(* IEC 61131-3 sources: PortalRobot/Portal_robot/Device/application, 34 files *)

(* ---- Persistent_Value.gvl.st ---- *)
{attribute 'qualified_only'}
VAR_GLOBAL PERSISTENT RETAIN
	// Постоянное хранилище базовых точек в энергонезависимой памяти контроллера.
	// Размер 15 сохранён ради совместимости со старой раскладкой: позиции 2, 6 и 10
	// (legacy MACHINE_x_INSIDE) больше не публикуются и не участвуют в готовности.
	astRetainPoints : ARRAY [1..GVL_POINT.iPersistentPointCapacity] OF ST_POINT;
	udiPointStorageVersion : UDINT;

	// Геометрический контроль: настройки, память станций и вызовы.
	astConfig : ARRAY [1..2] OF ST_GEOMETRY_CONFIG;
	astMemory : ARRAY [1..2] OF ST_GEOMETRY_MEMORY;
	astRetainCalls : ARRAY [1..3] OF ST_GEOMETRY_CALL;
	udiNextCallId : UDINT;
	udiEventSequence : UDINT;
	xAutoEnabled : BOOL := FALSE;
	auiPeriod : ARRAY [1..3] OF UINT := [20, 20, 20];
	auiCount : ARRAY [1..3] OF UINT;
	xWaitWhenOccupied : BOOL := TRUE;
	tTransportTimeout : TIME := T#10S;
	tDriveFeedbackTimeout : TIME := T#3S;
	tResetPulse : TIME := T#1S;
	tWaitWarningTimeout : TIME := T#180S; // Ожидание готовой вызванной детали в станке до WARNING

	// Постоянный шаг сетки для расчёта координат робота, отдельно по типам магазинов.
	lrStaticPitchX : LREAL := 60.0;
	lrStaticPitchY : LREAL := 60.0;
	lrTwinPitchX : LREAL := 70.0;
	lrTwinPitchY : LREAL := 70.0;

	// Базы ГК для SIMULATION сохраняются отдельно от реальных координат.
	astSimulationConfig : ARRAY [1..2] OF ST_GEOMETRY_CONFIG;

	// Добавлено в конце списка: прежние 15 баз и их версия сохраняют раскладку.
	astMagazineCalibration : ARRAY [1..2] OF ST_MAGAZINE_CALIBRATION;
END_VAR

(* ---- PLC_PRG.AppendIoEvent.st ---- *)
METHOD PRIVATE AppendIoEvent
VAR_INPUT
    usiDirection : USINT;
    uiIndex : UINT;
    usiKind : USINT;
    xOld : BOOL;
    xNew : BOOL;
END_VAR
VAR
    uiSlot : UINT;
    sEvent : STRING(96);
END_VAR

// --- BEGIN IMPLEMENTATION ---

IF NOT xIoSnapshotPublishing THEN
    GVL_HMI.udiIoJournalRevision := GVL_HMI.udiIoJournalRevision + UDINT#1;
END_IF;
// Переполнение Seq открывает новый FIFO; идентификаторы не повторяются внутри эпохи.
IF GVL_HMI.udiIoJournalSequence = UDINT#4294967295 THEN
    GVL_HMI.udiIoBootCounter := GVL_HMI.udiIoBootCounter + UDINT#1;
    IF GVL_HMI.udiIoBootCounter = UDINT#0 THEN GVL_HMI.udiIoBootCounter := UDINT#1; END_IF;
    GVL_HMI.udiIoJournalSequence := UDINT#0;
    GVL_HMI.uiIoJournalHead := UINT#0;
    GVL_HMI.uiIoJournalCount := UINT#0;
END_IF;
uiSlot := (GVL_HMI.uiIoJournalHead MOD UINT#100) + UINT#1;
GVL_HMI.udiIoJournalSequence := GVL_HMI.udiIoJournalSequence + UDINT#1;
astIoEvent[uiSlot].udiSequence := GVL_HMI.udiIoJournalSequence;
astIoEvent[uiSlot].uliTimeMs := uliIoClockMs;
astIoEvent[uiSlot].usiDirection := usiDirection;
astIoEvent[uiSlot].uiIndex := uiIndex;
astIoEvent[uiSlot].usiKind := usiKind;
astIoEvent[uiSlot].xOld := xOld;
astIoEvent[uiSlot].xNew := xNew;
// Строка кодируется только для изменившегося слота, не для всего FIFO на каждом скане.
sEvent := CONCAT(UDINT_TO_STRING(GVL_HMI.udiIoJournalSequence), ';');
sEvent := CONCAT(sEvent, ULINT_TO_STRING(uliIoClockMs));
sEvent := CONCAT(sEvent, ';'); sEvent := CONCAT(sEvent, USINT_TO_STRING(usiDirection));
sEvent := CONCAT(sEvent, ';'); sEvent := CONCAT(sEvent, UINT_TO_STRING(uiIndex));
sEvent := CONCAT(sEvent, ';'); sEvent := CONCAT(sEvent, USINT_TO_STRING(usiKind));
sEvent := CONCAT(sEvent, ';'); sEvent := CONCAT(sEvent, USINT_TO_STRING(BOOL_TO_USINT(xOld)));
sEvent := CONCAT(sEvent, ';'); sEvent := CONCAT(sEvent, USINT_TO_STRING(BOOL_TO_USINT(xNew)));
GVL_HMI.asIoJournal[uiSlot] := sEvent;
GVL_HMI.uiIoJournalHead := uiSlot;
GVL_HMI.uiIoJournalCount := MIN(UINT#100, GVL_HMI.uiIoJournalCount + UINT#1);
IF NOT xIoSnapshotPublishing THEN
    GVL_HMI.udiIoJournalRevision := GVL_HMI.udiIoJournalRevision + UDINT#1;
END_IF;

(* ---- PLC_PRG.ApplyIoOutputOverrides.st ---- *)
METHOD PRIVATE ApplyIoOutputOverrides

// --- BEGIN IMPLEMENTATION ---

// Прямой ручной режим владеет всеми DO. Штатные уровни остаются отдельно для возврата программе.
axIoAutoDo[1] := GVL_PHYSICAL_IO.xDoMachine1HatchClosed;
axIoAutoDo[2] := GVL_PHYSICAL_IO.xDoMachine1HatchUnLock;
axIoAutoDo[3] := GVL_PHYSICAL_IO.xDoMachine1ClampChuck;
axIoAutoDo[4] := GVL_PHYSICAL_IO.xDoMachine1UnclampChuck;
axIoAutoDo[5] := GVL_PHYSICAL_IO.xDoMachine1StartCycle;
axIoAutoDo[6] := GVL_PHYSICAL_IO.xDoMachine2HatchClosed;
axIoAutoDo[7] := GVL_PHYSICAL_IO.xDoMachine2HatchUnLock;
axIoAutoDo[8] := GVL_PHYSICAL_IO.xDoMachine2ClampChuck;
axIoAutoDo[9] := GVL_PHYSICAL_IO.xDoMachine2UnclampChuck;
axIoAutoDo[10] := GVL_PHYSICAL_IO.xDoMachine2StartCycle;
axIoAutoDo[11] := GVL_PHYSICAL_IO.xDoMachine3HatchClosed;
axIoAutoDo[12] := GVL_PHYSICAL_IO.xDoMachine3HatchUnLock;
axIoAutoDo[13] := GVL_PHYSICAL_IO.xDoMachine3ClampChuck;
axIoAutoDo[14] := GVL_PHYSICAL_IO.xDoMachine3UnclampChuck;
axIoAutoDo[15] := GVL_PHYSICAL_IO.xDoMachine3StartCycle;
axIoAutoDo[16] := GVL_PHYSICAL_IO.xDoGripper1Open;
axIoAutoDo[17] := GVL_PHYSICAL_IO.xDoGripper2Open;
axIoAutoDo[18] := GVL_PHYSICAL_IO.xDoRotateToDetail;
axIoAutoDo[19] := GVL_PHYSICAL_IO.xDoDoor1Unlock;
axIoAutoDo[20] := GVL_PHYSICAL_IO.xDoDoor2Unlock;
axIoAutoDo[21] := GVL_PHYSICAL_IO.xDoDoor3Unlock;
axIoAutoDo[22] := GVL_PHYSICAL_IO.xDoDoor4Unlock;
axIoAutoDo[23] := GVL_PHYSICAL_IO.xDoSafetyRelayReset;
axIoAutoDo[24] := GVL_PHYSICAL_IO.xDoSignalTowerGreenOutput;
axIoAutoDo[25] := GVL_PHYSICAL_IO.xDoSignalTowerAmberOutput;
axIoAutoDo[26] := GVL_PHYSICAL_IO.xDoSignalTowerRedOutput;
axIoAutoDo[27] := GVL_PHYSICAL_IO.xDoDoor1ButtonLamp;
axIoAutoDo[28] := GVL_PHYSICAL_IO.xDoDoor2ButtonLamp;
axIoAutoDo[29] := GVL_PHYSICAL_IO.xDoDoor3ButtonLamp;
axIoAutoDo[30] := GVL_PHYSICAL_IO.xDoDoor4ButtonLamp;
axIoAutoDo[31] := GVL_PHYSICAL_IO.xDoMagazine1LockIn;
axIoAutoDo[32] := GVL_PHYSICAL_IO.xDoMagazine1LockOut;
axIoAutoDo[33] := GVL_PHYSICAL_IO.xDoMagazine1StopIn;
axIoAutoDo[34] := GVL_PHYSICAL_IO.xDoMagazine1StopOut;
axIoAutoDo[35] := GVL_PHYSICAL_IO.xDoMagazine1LiftUp;
axIoAutoDo[36] := GVL_PHYSICAL_IO.xDoMagazine1LiftDown;
axIoAutoDo[37] := FALSE; // Удалённый сигнал; индекс журнала не переиспользовать.
axIoAutoDo[38] := FALSE; // Удалённый сигнал; индекс журнала не переиспользовать.
axIoAutoDo[39] := FALSE; // Удалённый сигнал; индекс журнала не переиспользовать.
axIoAutoDo[40] := GVL_PHYSICAL_IO.xDoCellAlarmHorn;
axIoAutoDo[41] := GVL_PHYSICAL_IO.xDoGk1DriveRun;
axIoAutoDo[42] := GVL_PHYSICAL_IO.xDoGk1DriveReset;
axIoAutoDo[43] := GVL_PHYSICAL_IO.xDoMagazine2LockIn;
axIoAutoDo[44] := GVL_PHYSICAL_IO.xDoMagazine2LockOut;
axIoAutoDo[45] := GVL_PHYSICAL_IO.xDoMagazine2StopIn;
axIoAutoDo[46] := GVL_PHYSICAL_IO.xDoMagazine2StopOut;
axIoAutoDo[47] := GVL_PHYSICAL_IO.xDoMagazine2LiftUp;
axIoAutoDo[48] := GVL_PHYSICAL_IO.xDoMagazine2LiftDown;
axIoAutoDo[49] := GVL_PHYSICAL_IO.xDoGk2DriveRun;
axIoAutoDo[50] := GVL_PHYSICAL_IO.xDoGk2DriveReset;
IF xIoManualActive AND NOT GVL_CELL_CONTROL.xManual THEN xIoManualActive := FALSE; END_IF;
GVL_HMI.xIoManualControlActive := xIoManualActive;
GVL_HMI.xIoDoOverrideAllowed := xIoManualActive AND GVL_CELL_CONTROL.xManual;
GVL_HMI.uiIoDoBlockReason := GVL_HMI.uiIoOverrideBlockReason;
IF GVL_HMI.xIoDoOverrideAllowed THEN GVL_HMI.uiIoDoBlockReason := UINT#0; END_IF;

FOR uiIoIndex := UINT#1 TO UINT#50 DO
    // 37..39 удалены из каталога; остальные индексы сохраняют смысл старых событий.
    IF (uiIoIndex >= UINT#37) AND (uiIoIndex <= UINT#39) THEN
        axIoDoForced[uiIoIndex] := FALSE;
        axIoDoForceValue[uiIoIndex] := FALSE;
    END_IF;
    axIoDoAllowed[uiIoIndex] := GVL_HMI.xIoDoOverrideAllowed AND ((uiIoIndex < UINT#37) OR (uiIoIndex > UINT#39));
    axIoDoOnAllowed[uiIoIndex] := axIoDoAllowed[uiIoIndex]; // Совместимость транспорта: включение и отключение равноправны.
    axIoDoInhibited[uiIoIndex] := FALSE; // Старый механизм блокировки снят.
    IF NOT xIoManualActive AND axIoDoForced[uiIoIndex] THEN
        IF xIoManualEndedByOperator THEN
            AppendIoEvent(usiDirection := USINT#2, uiIndex := uiIoIndex, usiKind := USINT#8,
                xOld := axIoDoForceValue[uiIoIndex], xNew := axIoAutoDo[uiIoIndex]);
        ELSE
            AppendIoEvent(usiDirection := USINT#2, uiIndex := uiIoIndex, usiKind := USINT#9,
                xOld := axIoDoForceValue[uiIoIndex], xNew := axIoAutoDo[uiIoIndex]);
        END_IF;
        axIoDoForced[uiIoIndex] := FALSE;
    END_IF;
END_FOR;

xIoDoRejected := FALSE;
udiIoRequestSeq := GVL_HMI.udiIoOverrideCommandSeq;
uiIoRequestAction := GVL_HMI.uiIoOverrideAction;
uiIoRequestIndex := GVL_HMI.uiIoOverrideIndex;
xIoRequestValue := GVL_HMI.xIoOverrideValue;
IF (udiIoRequestSeq <> GVL_HMI.udiIoOverrideAckSeq) AND (uiIoRequestAction >= UINT#4) AND (uiIoRequestAction <= UINT#9) THEN
    IF uiIoRequestAction <= UINT#6 THEN
        GVL_HMI.uiIoOverrideResult := UINT#3;
        IF NOT IsHmiCommandFresh(udiIssuedAtMs := GVL_HMI.udiIoOverrideIssuedAtMs) THEN
            GVL_HMI.uiIoOverrideResult := UINT#4;
        ELSIF uiIoRequestAction = UINT#6 THEN
            FOR uiIoIndex := UINT#1 TO UINT#50 DO
                IF axIoDoForced[uiIoIndex] THEN
                    AppendIoEvent(usiDirection := USINT#2, uiIndex := uiIoIndex, usiKind := USINT#8,
                        xOld := axIoDoForceValue[uiIoIndex], xNew := axIoAutoDo[uiIoIndex]);
                END_IF;
                axIoDoForceValue[uiIoIndex] := axIoAutoDo[uiIoIndex];
                axIoDoForced[uiIoIndex] := FALSE;
            END_FOR;
            GVL_HMI.uiIoOverrideResult := UINT#1;
        ELSIF (uiIoRequestIndex >= UINT#1) AND (uiIoRequestIndex <= UINT#50) AND ((uiIoRequestIndex < UINT#37) OR (uiIoRequestIndex > UINT#39)) THEN
            IF uiIoRequestAction = UINT#5 THEN
                IF axIoDoForced[uiIoRequestIndex] THEN
                    AppendIoEvent(usiDirection := USINT#2, uiIndex := uiIoRequestIndex, usiKind := USINT#8,
                        xOld := axIoDoForceValue[uiIoRequestIndex], xNew := axIoAutoDo[uiIoRequestIndex]);
                END_IF;
                axIoDoForceValue[uiIoRequestIndex] := axIoAutoDo[uiIoRequestIndex];
                axIoDoForced[uiIoRequestIndex] := FALSE;
                GVL_HMI.uiIoOverrideResult := UINT#1;
            ELSIF GVL_HMI.xIoDoOverrideAllowed THEN
                IF NOT axIoDoForced[uiIoRequestIndex] OR (axIoDoForceValue[uiIoRequestIndex] <> xIoRequestValue) THEN
                    AppendIoEvent(usiDirection := USINT#2, uiIndex := uiIoRequestIndex, usiKind := USINT#7,
                        xOld := axIoOutput[uiIoRequestIndex], xNew := xIoRequestValue);
                END_IF;
                axIoDoForced[uiIoRequestIndex] := TRUE;
                axIoDoForceValue[uiIoRequestIndex] := xIoRequestValue;
                IF (uiIoRequestIndex >= UINT#31) AND (uiIoRequestIndex <= UINT#36) THEN axIoMagazineInvalidated[1] := TRUE;
                ELSIF (uiIoRequestIndex >= UINT#43) AND (uiIoRequestIndex <= UINT#48) THEN axIoMagazineInvalidated[2] := TRUE;
                END_IF;
                GVL_HMI.uiIoOverrideResult := UINT#1;
            ELSE
                GVL_HMI.uiIoOverrideResult := UINT#2;
            END_IF;
        END_IF;
    END_IF;
    xIoDoRejected := GVL_HMI.uiIoOverrideResult <> UINT#1;
    GVL_HMI.udiIoOverrideAckSeq := udiIoRequestSeq;
END_IF;

// Намеренно без Safety, пар катушек, режима Modbus, импульсных ограничений и технологических FB.
IF xIoManualActive THEN
    GVL_PHYSICAL_IO.xDoMachine1HatchClosed := axIoDoForceValue[1];
    GVL_PHYSICAL_IO.xDoMachine1HatchUnLock := axIoDoForceValue[2];
    GVL_PHYSICAL_IO.xDoMachine1ClampChuck := axIoDoForceValue[3];
    GVL_PHYSICAL_IO.xDoMachine1UnclampChuck := axIoDoForceValue[4];
    GVL_PHYSICAL_IO.xDoMachine1StartCycle := axIoDoForceValue[5];
    GVL_PHYSICAL_IO.xDoMachine2HatchClosed := axIoDoForceValue[6];
    GVL_PHYSICAL_IO.xDoMachine2HatchUnLock := axIoDoForceValue[7];
    GVL_PHYSICAL_IO.xDoMachine2ClampChuck := axIoDoForceValue[8];
    GVL_PHYSICAL_IO.xDoMachine2UnclampChuck := axIoDoForceValue[9];
    GVL_PHYSICAL_IO.xDoMachine2StartCycle := axIoDoForceValue[10];
    GVL_PHYSICAL_IO.xDoMachine3HatchClosed := axIoDoForceValue[11];
    GVL_PHYSICAL_IO.xDoMachine3HatchUnLock := axIoDoForceValue[12];
    GVL_PHYSICAL_IO.xDoMachine3ClampChuck := axIoDoForceValue[13];
    GVL_PHYSICAL_IO.xDoMachine3UnclampChuck := axIoDoForceValue[14];
    GVL_PHYSICAL_IO.xDoMachine3StartCycle := axIoDoForceValue[15];
    GVL_PHYSICAL_IO.xDoGripper1Open := axIoDoForceValue[16];
    GVL_PHYSICAL_IO.xDoGripper2Open := axIoDoForceValue[17];
    GVL_PHYSICAL_IO.xDoRotateToDetail := axIoDoForceValue[18];
    GVL_PHYSICAL_IO.xDoDoor1Unlock := axIoDoForceValue[19];
    GVL_PHYSICAL_IO.xDoDoor2Unlock := axIoDoForceValue[20];
    GVL_PHYSICAL_IO.xDoDoor3Unlock := axIoDoForceValue[21];
    GVL_PHYSICAL_IO.xDoDoor4Unlock := axIoDoForceValue[22];
    GVL_PHYSICAL_IO.xDoSafetyRelayReset := axIoDoForceValue[23];
    GVL_PHYSICAL_IO.xDoSignalTowerGreenOutput := axIoDoForceValue[24];
    GVL_PHYSICAL_IO.xDoSignalTowerAmberOutput := axIoDoForceValue[25];
    GVL_PHYSICAL_IO.xDoSignalTowerRedOutput := axIoDoForceValue[26];
    GVL_PHYSICAL_IO.xDoDoor1ButtonLamp := axIoDoForceValue[27];
    GVL_PHYSICAL_IO.xDoDoor2ButtonLamp := axIoDoForceValue[28];
    GVL_PHYSICAL_IO.xDoDoor3ButtonLamp := axIoDoForceValue[29];
    GVL_PHYSICAL_IO.xDoDoor4ButtonLamp := axIoDoForceValue[30];
    GVL_PHYSICAL_IO.xDoMagazine1LockIn := axIoDoForceValue[31];
    GVL_PHYSICAL_IO.xDoMagazine1LockOut := axIoDoForceValue[32];
    GVL_PHYSICAL_IO.xDoMagazine1StopIn := axIoDoForceValue[33];
    GVL_PHYSICAL_IO.xDoMagazine1StopOut := axIoDoForceValue[34];
    GVL_PHYSICAL_IO.xDoMagazine1LiftUp := axIoDoForceValue[35];
    GVL_PHYSICAL_IO.xDoMagazine1LiftDown := axIoDoForceValue[36];
    GVL_PHYSICAL_IO.xDoCellAlarmHorn := axIoDoForceValue[40];
    GVL_PHYSICAL_IO.xDoGk1DriveRun := axIoDoForceValue[41];
    GVL_PHYSICAL_IO.xDoGk1DriveReset := axIoDoForceValue[42];
    GVL_PHYSICAL_IO.xDoMagazine2LockIn := axIoDoForceValue[43];
    GVL_PHYSICAL_IO.xDoMagazine2LockOut := axIoDoForceValue[44];
    GVL_PHYSICAL_IO.xDoMagazine2StopIn := axIoDoForceValue[45];
    GVL_PHYSICAL_IO.xDoMagazine2StopOut := axIoDoForceValue[46];
    GVL_PHYSICAL_IO.xDoMagazine2LiftUp := axIoDoForceValue[47];
    GVL_PHYSICAL_IO.xDoMagazine2LiftDown := axIoDoForceValue[48];
    GVL_PHYSICAL_IO.xDoGk2DriveRun := axIoDoForceValue[49];
    GVL_PHYSICAL_IO.xDoGk2DriveReset := axIoDoForceValue[50];
END_IF;

(* ---- PLC_PRG.BuildRobotResetDependencies.st ---- *)
METHOD PRIVATE BuildRobotResetDependencies
VAR
	uiOwner : UINT;
	dwOwnerBit : DWORD;
END_VAR

// --- BEGIN IMPLEMENTATION ---

// Снимок после вызовов владельцев, перед FB_ROBOT. Не смешиваем первичную
// причину оборудования с зависимой ошибкой родителя и не изменяем GVL-теги.
stRobotResetDependencies.dwStopOwners := DWORD#0;
stRobotResetDependencies.dwLiveCauses := DWORD#0;
stRobotResetDependencies.dwResetBusy := DWORD#0;
FOR uiOwner := UINT#1 TO UINT#3 DO
	dwOwnerBit := SHL(DWORD#1, uiOwner - UINT#1);
	IF GVL_MACHINE.Status[uiOwner].xCriticalError THEN
		stRobotResetDependencies.dwStopOwners := stRobotResetDependencies.dwStopOwners OR dwOwnerBit;
		IF GVL_MACHINE.Status[uiOwner].stIo.xAlarm THEN
			stRobotResetDependencies.dwLiveCauses := stRobotResetDependencies.dwLiveCauses OR dwOwnerBit;
		END_IF;
	END_IF;
END_FOR;
FOR uiOwner := UINT#1 TO UINT#2 DO
	dwOwnerBit := SHL(DWORD#1, uiOwner + UINT#2);
	IF GVL_MAGAZINE.astPartStatus[uiOwner].xRobotStopRequired THEN
		stRobotResetDependencies.dwStopOwners := stRobotResetDependencies.dwStopOwners OR dwOwnerBit;
	END_IF;
	dwOwnerBit := SHL(DWORD#1, uiOwner + UINT#4);
	IF GVL_GEOMETRY_CONTROL.xSupported AND GVL_GEOMETRY_CONTROL.astStatus[uiOwner].xRobotStopRequired THEN
		stRobotResetDependencies.dwStopOwners := stRobotResetDependencies.dwStopOwners OR dwOwnerBit;
		IF GEOMETRY[uiOwner].xDriveAlarm THEN
			stRobotResetDependencies.dwLiveCauses := stRobotResetDependencies.dwLiveCauses OR dwOwnerBit;
		END_IF;
	END_IF;
	IF GVL_GEOMETRY_CONTROL.xSupported AND GVL_GEOMETRY_CONTROL.astStatus[uiOwner].xResetBusy THEN
		stRobotResetDependencies.dwResetBusy := stRobotResetDependencies.dwResetBusy OR dwOwnerBit;
	END_IF;
	dwOwnerBit := SHL(DWORD#1, uiOwner + UINT#6);
	IF (GVL_TWO_PALLET.uiMode = UINT#1) AND axTwinRobotStopLatched[uiOwner] THEN
		stRobotResetDependencies.dwStopOwners := stRobotResetDependencies.dwStopOwners OR dwOwnerBit;
		IF TWIN[uiOwner].Input.xDriveError THEN
			stRobotResetDependencies.dwLiveCauses := stRobotResetDependencies.dwLiveCauses OR dwOwnerBit;
		END_IF;
	END_IF;
END_FOR;

(* ---- PLC_PRG.InvalidateMagazineCalibration.st ---- *)
METHOD PRIVATE InvalidateMagazineCalibration
VAR_INPUT
	uiMagazine : UINT;
END_VAR
VAR
	eOrigin : E_POINT_NAME;
	ePointB : E_POINT_NAME;
	ePointC : E_POINT_NAME;
END_VAR

// --- BEGIN IMPLEMENTATION ---

// Все три признака снимаются одной PLC-транзакцией; координаты остаются черновиком.
IF (uiMagazine >= UINT#1) AND (uiMagazine <= UINT#2) THEN
	IF uiMagazine = UINT#1 THEN
		eOrigin := E_POINT_NAME.MAGAZINE_1_DETAIL;
		ePointB := E_POINT_NAME.MAGAZINE_1_AXIS_X;
		ePointC := E_POINT_NAME.MAGAZINE_1_AXIS_Y;
	ELSE
		eOrigin := E_POINT_NAME.MAGAZINE_2_DETAIL;
		ePointB := E_POINT_NAME.MAGAZINE_2_AXIS_X;
		ePointC := E_POINT_NAME.MAGAZINE_2_AXIS_Y;
	END_IF;
	Persistent_Value.astRetainPoints[UINT#13 + uiMagazine].xConfigured := FALSE;
	Persistent_Value.astMagazineCalibration[uiMagazine].astReference[1].xConfigured := FALSE;
	Persistent_Value.astMagazineCalibration[uiMagazine].astReference[2].xConfigured := FALSE;
	GVL_POINT.Points[eOrigin].xConfigured := FALSE;
	GVL_POINT.Points[ePointB].xConfigured := FALSE;
	GVL_POINT.Points[ePointC].xConfigured := FALSE;
	axMagazinePointsReady[uiMagazine] := FALSE;
	astMagazineFrame[uiMagazine].xReady := FALSE;
	GVL_HMI.astMagazineCalibrationStatus[uiMagazine].xReady := FALSE;
	xPointTableReady := FALSE;
END_IF;

(* ---- PLC_PRG.IsHmiCommandFresh.st ---- *)
METHOD PRIVATE IsHmiCommandFresh : BOOL
VAR_INPUT
	udiIssuedAtMs : UDINT;
END_VAR
VAR
	uliAgeMs : ULINT;
END_VAR

// --- BEGIN IMPLEMENTATION ---

// Explicit modulo-2^32 age: TIME() rolls over after about 49 days.
IF udiHmiCommandNowMs >= udiIssuedAtMs THEN
	uliAgeMs := UDINT_TO_ULINT(udiHmiCommandNowMs) - UDINT_TO_ULINT(udiIssuedAtMs);
ELSE
	uliAgeMs := ULINT#4294967296 + UDINT_TO_ULINT(udiHmiCommandNowMs) - UDINT_TO_ULINT(udiIssuedAtMs);
END_IF;
IsHmiCommandFresh := uliAgeMs <= UDINT_TO_ULINT(
	TIME_TO_UDINT(GVL_CELL_SETTINGS.tHmiCommandFreshnessTimeout)
);

(* ---- PLC_PRG.PublishGeometryControl.st ---- *)
METHOD PRIVATE PublishGeometryControl
VAR
	uiWarningEvent : UINT;
END_VAR

// --- BEGIN IMPLEMENTATION ---

GVL_HMI.astGeometryStatus := GVL_GEOMETRY_CONTROL.astStatus;
// Подсветка следует накопленному предупреждению, включая его сброс в этом скане.
IF ALARM_MANAGER.xEventsUpdated OR NOT xHmiTablesInitialized THEN
xGeometryWaitWarningActive := FALSE;
FOR uiWarningEvent := UINT#1 TO UINT#100 DO
	IF GVL_ALARM.Events[uiWarningEvent].xActive
	AND (GVL_ALARM.Events[uiWarningEvent].eSource = E_ALARM_SOURCE.CELL)
	AND (GVL_ALARM.Events[uiWarningEvent].eSeverity = E_ALARM_SEVERITY.WARNING)
	AND (GVL_ALARM.Events[uiWarningEvent].uiCode = UINT#52) THEN xGeometryWaitWarningActive := TRUE; END_IF;
END_FOR;
END_IF;
FOR uiGeometry := UINT#1 TO UINT#2 DO
	GVL_HMI.astGeometryStatus[uiGeometry].xCallWaitWarning := xGeometryWaitWarningActive
		AND (GVL_GEOMETRY_CONTROL.astStatus[uiGeometry].xEnabled
			OR NOT (GVL_GEOMETRY_CONTROL.astStatus[1].xEnabled OR GVL_GEOMETRY_CONTROL.astStatus[2].xEnabled));
END_FOR;
GVL_HMI.astGeometryConfig := GVL_GEOMETRY_CONTROL.astActiveConfig;
GVL_HMI.astGeometryCalls := GVL_GEOMETRY_CONTROL.astCalls;
GVL_HMI.auiGeometryPeriod := Persistent_Value.auiPeriod;
GVL_HMI.auiGeometryCount := GVL_GEOMETRY_CONTROL.auiActiveCount;
GVL_HMI.axGeometryCallAllowed := GVL_GEOMETRY_CONTROL.axCallAllowed;
GVL_HMI.axGeometryCancelAllowed := GVL_GEOMETRY_CONTROL.axCancelAllowed;
GVL_HMI.xGeometryAutoEnabled := Persistent_Value.xAutoEnabled;
GVL_HMI.xGeometryAutoChangeAllowed := GVL_GEOMETRY_CONTROL.xAutoChangeAllowed;
GVL_HMI.xGeometrySupported := GVL_GEOMETRY_CONTROL.xSupported;
GVL_HMI.xGeometryWaitWhenOccupied := Persistent_Value.xWaitWhenOccupied;
GVL_HMI.tGeometryTransportTimeout := Persistent_Value.tTransportTimeout;
GVL_HMI.tGeometryFeedbackTimeout := Persistent_Value.tDriveFeedbackTimeout;
GVL_HMI.tGeometryResetPulse := Persistent_Value.tResetPulse;
GVL_HMI.tGeometryWaitWarningTimeout := Persistent_Value.tWaitWarningTimeout;
GVL_HMI.xGeometrySettingsAllowed := GVL_GEOMETRY_CONTROL.xSettingsAllowed;
// Снимок FIFO имеет версию: gateway читает одинаковый Seq до/после payload.
IF NOT xHmiTablesInitialized
OR (GVL_HMI.udiGeometryEventSequence <> Persistent_Value.udiEventSequence) THEN
    GVL_HMI.udiGeometryEventSequence := UDINT#0;
    GVL_HMI.astGeometryEvents := GVL_GEOMETRY_CONTROL.astEvents;
    GVL_HMI.udiGeometryEventSequence := Persistent_Value.udiEventSequence;
END_IF;
IF GVL_CELL_SETTINGS.eTestEnvironment = E_CELL_TEST_ENVIRONMENT.NORMAL THEN
	Persistent_Value.astMemory := GVL_GEOMETRY_CONTROL.astActiveMemory;
	Persistent_Value.astRetainCalls := GVL_GEOMETRY_CONTROL.astCalls;
	Persistent_Value.auiCount := GVL_GEOMETRY_CONTROL.auiActiveCount;
ELSE
	GVL_GEOMETRY_CONTROL.astSimulationMemory := GVL_GEOMETRY_CONTROL.astActiveMemory;
	GVL_GEOMETRY_CONTROL.astSimulationCalls := GVL_GEOMETRY_CONTROL.astCalls;
	GVL_GEOMETRY_CONTROL.auiSimulationCount := GVL_GEOMETRY_CONTROL.auiActiveCount;
END_IF;
// Фиксированные владельцы счётчиков: переключение среды не меняет идентичность
// OPC UA тега и не превращает старое значение NORMAL в выпуск SIMULATION.
FOR uiGeometry := UINT#1 TO UINT#2 DO
	GVL_HMI.audiGeometryProducedNormal[uiGeometry] := Persistent_Value.astMemory[uiGeometry].udiProducedPartsTotal;
	GVL_HMI.audiGeometryProducedSimulation[uiGeometry] := GVL_GEOMETRY_CONTROL.astSimulationMemory[uiGeometry].udiProducedPartsTotal;
END_FOR;

(* ---- PLC_PRG.PublishHmi.st ---- *)
METHOD PRIVATE PublishHmi

// --- BEGIN IMPLEMENTATION ---

// Единый снимок состояния для внешней визуализации.
GVL_HMI.udiPlcHeartbeat := GVL_HMI.udiPlcHeartbeat + 1;
GVL_HMI.xHmiConnectionAlive := xHmiConnectionAlive;
GVL_HMI.xManualRecoveryActive := xManualRecoveryActive;
GVL_HMI.xGlobalError := GVL_CELL_CONTROL.xGlobalError;
GVL_HMI.xCellManual := GVL_CELL_CONTROL.xManual;
// Отказ тоже потребляет транзакцию: она не исполнится позже сама собой.
GVL_HMI.udiCellModeAckSeq := udiCellModeCommandSnapshot;
GVL_HMI.xErrorSimulationEnabled := GVL_CELL_SETTINGS.xErrorSimulationEnabled;
GVL_HMI.stSafetyFaultStatus := CELL_SAFETY.FaultStatus;
GVL_HMI.xSimulationAccelerationActive := GVL_CELL_SETTINGS.xSimulationAccelerationActive;
GVL_HMI.xSimulationAccelerationChangeAllowed := GVL_CELL_SETTINGS.xSimulationAccelerationChangeAllowed;
GVL_HMI.uiSimulationTimeFactorApplied := GVL_CELL_SETTINGS.uiSimulationTimeFactorApplied;
GVL_HMI.xSimulationAccelerationPending := GVL_CELL_SETTINGS.xSimulationAccelerationPending;
GVL_HMI.xSimulationAccelerationBusy := GVL_CELL_SETTINGS.xSimulationAccelerationBusy;
GVL_HMI.xSimulationAccelerationError := GVL_CELL_SETTINGS.xSimulationAccelerationError;
GVL_HMI.udiSimulationAccelerationErrorId := GVL_CELL_SETTINGS.udiSimulationAccelerationErrorId;
GVL_HMI.lrSafetyHomeX := GVL_POINT.Points[E_POINT_NAME.HOME_SAFETY].X;
GVL_HMI.lrSafetyHomeY := GVL_POINT.Points[E_POINT_NAME.HOME_SAFETY].Y;
GVL_HMI.lrSafetyHomeZ := GVL_POINT.Points[E_POINT_NAME.HOME_SAFETY].Z;
GVL_HMI.lrSafetyHomeSpeedFactor := GVL_POINT.Points[E_POINT_NAME.HOME_SAFETY].SpeedFactor;
GVL_HMI.lrSafetyHomeToleranceX := GVL_CELL_SETTINGS.lrSafetyHomeToleranceX;
GVL_HMI.lrSafetyHomeToleranceY := GVL_CELL_SETTINGS.lrSafetyHomeToleranceY;
GVL_HMI.lrSafetyHomeToleranceZ := GVL_CELL_SETTINGS.lrSafetyHomeToleranceZ;
GVL_HMI.rRobotAccelerationPercent := GVL_CELL_SETTINGS.rRobotAccelerationPercent;
GVL_HMI.rRobotDecelerationPercent := GVL_CELL_SETTINGS.rRobotDecelerationPercent;
GVL_HMI.rRobotJerkPercent := GVL_CELL_SETTINGS.rRobotJerkPercent;
GVL_HMI.lrRobotHaltDeceleration := GVL_CELL_SETTINGS.lrRobotHaltDeceleration;
GVL_HMI.lrRobotHaltJerk := GVL_CELL_SETTINGS.lrRobotHaltJerk;
GVL_HMI.stCellMachineTimeouts := GVL_CELL_SETTINGS.stMachineTimeouts;
GVL_HMI.stCellAxisTimeouts := GVL_CELL_SETTINGS.stAxisTimeouts;
GVL_HMI.stCellAxisGroupTimeouts := GVL_CELL_SETTINGS.stAxisGroupTimeouts;
GVL_HMI.tPointCheckStartTimeout := GVL_CELL_SETTINGS.tPointCheckStartTimeout;
GVL_HMI.tSimulationDynamicsTimeout := GVL_CELL_SETTINGS.tSimulationDynamicsTimeout;
GVL_HMI.tHmiWatchdogTimeout := GVL_CELL_SETTINGS.tHmiWatchdogTimeout;
GVL_HMI.tMobileMotionWatchdogTimeout := GVL_CELL_SETTINGS.tMobileMotionWatchdogTimeout;
GVL_HMI.tPointCheckWatchdogTimeout := GVL_CELL_SETTINGS.tPointCheckWatchdogTimeout;
GVL_HMI.tHmiCommandFreshnessTimeout := GVL_CELL_SETTINGS.tHmiCommandFreshnessTimeout;
GVL_HMI.tAlarmHornDuration := GVL_CELL_SETTINGS.tAlarmHornDuration;
GVL_HMI.tInputFilterRise := GVL_CELL_SETTINGS.tInputFilterRise;
GVL_HMI.tInputFilterFall := GVL_CELL_SETTINGS.tInputFilterFall;
GVL_HMI.xIoFilterSettingsChangeAllowed := GVL_CELL_SETTINGS.xIoFilterSettingsChangeAllowed;
GVL_HMI.xPhysicalIoActive := GVL_PHYSICAL_IO.xNormalActive
	AND (GVL_CELL_SETTINGS.eTestEnvironment = E_CELL_TEST_ENVIRONMENT.NORMAL);
GVL_HMI.xPhysicalIoMappingVerified := GVL_PHYSICAL_IO.xMappingVerified;
GVL_HMI.xCellSettingsChangeAllowed := GVL_CELL_SETTINGS.xCellSettingsChangeAllowed;
GVL_HMI.rPointCheckSpeedPercent := GVL_CELL_SETTINGS.rPointCheckSpeedPercent;
GVL_HMI.xPointCheckActive := xPointCheckActive;
IF xPointCheckActive THEN
	GVL_HMI.rPointCheckAppliedSpeedPercent := rPointCheckLatchedSpeed;
ELSE
	GVL_HMI.rPointCheckAppliedSpeedPercent := GVL_CELL_SETTINGS.rPointCheckSpeedPercent;
END_IF;
GVL_HMI.xPointTableReady := xPointTableReady;
GVL_HMI.astPointEditorPoints[1] := GVL_POINT.Points[E_POINT_NAME.MACHINE_1_ABOVE];
GVL_HMI.astPointEditorPoints[2] := GVL_POINT.Points[E_POINT_NAME.MACHINE_1_CHUCK_APROACH];
GVL_HMI.astPointEditorPoints[3] := GVL_POINT.Points[E_POINT_NAME.MACHINE_1_CHUCK_POSITION];
GVL_HMI.astPointEditorPoints[4] := GVL_POINT.Points[E_POINT_NAME.MACHINE_2_ABOVE];
GVL_HMI.astPointEditorPoints[5] := GVL_POINT.Points[E_POINT_NAME.MACHINE_2_CHUCK_APROACH];
GVL_HMI.astPointEditorPoints[6] := GVL_POINT.Points[E_POINT_NAME.MACHINE_2_CHUCK_POSITION];
GVL_HMI.astPointEditorPoints[7] := GVL_POINT.Points[E_POINT_NAME.MACHINE_3_ABOVE];
GVL_HMI.astPointEditorPoints[8] := GVL_POINT.Points[E_POINT_NAME.MACHINE_3_CHUCK_APROACH];
GVL_HMI.astPointEditorPoints[9] := GVL_POINT.Points[E_POINT_NAME.MACHINE_3_CHUCK_POSITION];
GVL_HMI.astPointEditorPoints[10] := GVL_POINT.Points[E_POINT_NAME.HOME_SAFETY];
GVL_HMI.astPointEditorPoints[11] := GVL_POINT.Points[E_POINT_NAME.MAGAZINE_1_DETAIL];
GVL_HMI.astPointEditorPoints[12] := GVL_POINT.Points[E_POINT_NAME.MAGAZINE_2_DETAIL];
GVL_HMI.astPointEditorPoints[13] := GVL_POINT.Points[E_POINT_NAME.GEOMETRY_1_PLACE];
GVL_HMI.astPointEditorPoints[14] := GVL_POINT.Points[E_POINT_NAME.GEOMETRY_2_PLACE];
GVL_HMI.astPointEditorPoints[15] := GVL_POINT.Points[E_POINT_NAME.MAGAZINE_1_AXIS_X];
GVL_HMI.astPointEditorPoints[16] := GVL_POINT.Points[E_POINT_NAME.MAGAZINE_1_AXIS_Y];
GVL_HMI.astPointEditorPoints[17] := GVL_POINT.Points[E_POINT_NAME.MAGAZINE_2_AXIS_X];
GVL_HMI.astPointEditorPoints[18] := GVL_POINT.Points[E_POINT_NAME.MAGAZINE_2_AXIS_Y];
GVL_HMI.auiPointEditorPointId[1] := TO_UINT(E_POINT_NAME.MACHINE_1_ABOVE);
GVL_HMI.auiPointEditorPointId[2] := TO_UINT(E_POINT_NAME.MACHINE_1_CHUCK_APROACH);
GVL_HMI.auiPointEditorPointId[3] := TO_UINT(E_POINT_NAME.MACHINE_1_CHUCK_POSITION);
GVL_HMI.auiPointEditorPointId[4] := TO_UINT(E_POINT_NAME.MACHINE_2_ABOVE);
GVL_HMI.auiPointEditorPointId[5] := TO_UINT(E_POINT_NAME.MACHINE_2_CHUCK_APROACH);
GVL_HMI.auiPointEditorPointId[6] := TO_UINT(E_POINT_NAME.MACHINE_2_CHUCK_POSITION);
GVL_HMI.auiPointEditorPointId[7] := TO_UINT(E_POINT_NAME.MACHINE_3_ABOVE);
GVL_HMI.auiPointEditorPointId[8] := TO_UINT(E_POINT_NAME.MACHINE_3_CHUCK_APROACH);
GVL_HMI.auiPointEditorPointId[9] := TO_UINT(E_POINT_NAME.MACHINE_3_CHUCK_POSITION);
GVL_HMI.auiPointEditorPointId[10] := TO_UINT(E_POINT_NAME.HOME_SAFETY);
GVL_HMI.auiPointEditorPointId[11] := TO_UINT(E_POINT_NAME.MAGAZINE_1_DETAIL);
GVL_HMI.auiPointEditorPointId[12] := TO_UINT(E_POINT_NAME.MAGAZINE_2_DETAIL);
GVL_HMI.auiPointEditorPointId[13] := TO_UINT(E_POINT_NAME.GEOMETRY_1_PLACE);
GVL_HMI.auiPointEditorPointId[14] := TO_UINT(E_POINT_NAME.GEOMETRY_2_PLACE);
GVL_HMI.auiPointEditorPointId[15] := TO_UINT(E_POINT_NAME.MAGAZINE_1_AXIS_X);
GVL_HMI.auiPointEditorPointId[16] := TO_UINT(E_POINT_NAME.MAGAZINE_1_AXIS_Y);
GVL_HMI.auiPointEditorPointId[17] := TO_UINT(E_POINT_NAME.MAGAZINE_2_AXIS_X);
GVL_HMI.auiPointEditorPointId[18] := TO_UINT(E_POINT_NAME.MAGAZINE_2_AXIS_Y);
GVL_HMI.astMagazineCalibrationStatus[1].astPoints[1] := GVL_POINT.Points[E_POINT_NAME.MAGAZINE_1_DETAIL];
GVL_HMI.astMagazineCalibrationStatus[1].astPoints[2] := GVL_POINT.Points[E_POINT_NAME.MAGAZINE_1_AXIS_X];
GVL_HMI.astMagazineCalibrationStatus[1].astPoints[3] := GVL_POINT.Points[E_POINT_NAME.MAGAZINE_1_AXIS_Y];
GVL_HMI.astMagazineCalibrationStatus[2].astPoints[1] := GVL_POINT.Points[E_POINT_NAME.MAGAZINE_2_DETAIL];
GVL_HMI.astMagazineCalibrationStatus[2].astPoints[2] := GVL_POINT.Points[E_POINT_NAME.MAGAZINE_2_AXIS_X];
GVL_HMI.astMagazineCalibrationStatus[2].astPoints[3] := GVL_POINT.Points[E_POINT_NAME.MAGAZINE_2_AXIS_Y];
// Метод публикуется после опор: новый режим не сопровождается прежними флагами A/B/C.
GVL_HMI.astMagazineCalibrationStatus[1].uiMethod := Persistent_Value.astMagazineCalibration[1].uiMethod;
GVL_HMI.astMagazineCalibrationStatus[2].uiMethod := Persistent_Value.astMagazineCalibration[2].uiMethod;
GVL_HMI.xModbusMode := GVL_ROBOT_MODBUS.xModeActive;
GVL_HMI.xRobotModeChangeAllowed := GVL_ROBOT_MODBUS.xRobotModeChangeAllowed;
GVL_HMI.xModbusSettingsChangeAllowed := GVL_ROBOT_MODBUS.xSettingsChangeAllowed;
GVL_HMI.stRobotModbusStatus := GVL_ROBOT_MODBUS.Status;
uiMagazine := GVL_CELL_MANAGER.Status.uiActiveMagazine;
IF (uiMagazine < UINT#1) OR (uiMagazine > UINT#2) THEN
	uiMagazine := UINT#1;
END_IF;
GVL_HMI.stTestObservability.uiSchemaVersion := UINT#3;
GVL_HMI.stTestObservability.uiReturnMagazine := CELL_MANAGER.uiReturnMagazine;
GVL_HMI.stTestObservability.udiAppliedScenarioSeq := GVL_HMI.udiTestScenarioAckSeq;
GVL_HMI.stTestObservability.uiCellState := TO_UINT(GVL_CELL_MANAGER.Diag.eState);
GVL_HMI.stTestObservability.uiRobotState := TO_UINT(GVL_ROBOT.Diag.eState);
GVL_HMI.stTestObservability.uiRobotAction := TO_UINT(GVL_ROBOT.Diag.eActiveAction);
GVL_HMI.stTestObservability.uiRobotPoint := TO_UINT(GVL_ROBOT.Diag.eActivePoint);
GVL_HMI.stTestObservability.uiActiveMagazine := GVL_CELL_MANAGER.Status.uiActiveMagazine;
GVL_HMI.stTestObservability.uiMagazineState := TO_UINT(GVL_MAGAZINE.astDiag[uiMagazine].eState);
GVL_HMI.stTestObservability.uiMagazineOperation := TO_UINT(GVL_MAGAZINE.astStatus[uiMagazine].eActualOperation);
GVL_HMI.stTestObservability.uiTakeSlot := SINT_TO_UINT(GVL_MAGAZINE.astStatus[uiMagazine].iSelectedBlank);
GVL_HMI.stTestObservability.uiPutSlot := SINT_TO_UINT(GVL_MAGAZINE.astStatus[uiMagazine].iSelectedFreeSlot);
GVL_HMI.stTestObservability.uiSelectedMachine := GVL_CELL_MANAGER.Status.uiSelectedMachine;
GVL_HMI.stTestObservability.uiSelectedType := GVL_MULTI_TYPE.CycleStatus.uiSelectedType;
GVL_HMI.stTestObservability.uiErrorSource := UINT#0;
GVL_HMI.stTestObservability.dwErrorCode := DWORD#0;
FOR uiMachine := 1 TO 3 DO
	GVL_HMI.stTestObservability.auiMachineState[uiMachine] := TO_UINT(GVL_MACHINE.Diag[uiMachine].eState);
	GVL_HMI.stTestObservability.auiMachineOperation[uiMachine] := TO_UINT(GVL_MACHINE.Diag[uiMachine].eActualOperation);
END_FOR;
IF GVL_ROBOT.Error.dwErrorActive <> DWORD#0 THEN
	GVL_HMI.stTestObservability.uiErrorSource := UINT#2;
	GVL_HMI.stTestObservability.dwErrorCode := GVL_ROBOT.Error.dwErrorActive;
ELSIF GVL_MAGAZINE.astError[1].dwErrorActive <> DWORD#0 THEN
	GVL_HMI.stTestObservability.uiErrorSource := UINT#3;
GVL_HMI.stTestObservability.dwErrorCode := GVL_MAGAZINE.astError[1].dwErrorActive;
ELSIF GVL_MAGAZINE.astError[2].dwErrorActive <> DWORD#0 THEN
	GVL_HMI.stTestObservability.uiErrorSource := UINT#7;
	GVL_HMI.stTestObservability.dwErrorCode := GVL_MAGAZINE.astError[2].dwErrorActive;
ELSIF GVL_CELL_MANAGER.Error.dwErrorActive <> DWORD#0 THEN
	GVL_HMI.stTestObservability.uiErrorSource := UINT#1;
	GVL_HMI.stTestObservability.dwErrorCode := GVL_CELL_MANAGER.Error.dwErrorActive;
ELSE
	FOR uiMachine := 1 TO 3 DO
		IF GVL_MACHINE.Error[uiMachine].dwErrorActive <> DWORD#0 THEN
			GVL_HMI.stTestObservability.uiErrorSource := uiMachine + UINT#3;
			GVL_HMI.stTestObservability.dwErrorCode := GVL_MACHINE.Error[uiMachine].dwErrorActive;
		END_IF;
	END_FOR;
END_IF;
FOR uiMachine := 1 TO 9 DO
	GVL_HMI.auiRobotModbusWriteRegisters[uiMachine] :=
		GVL_ROBOT_MODBUS.auiWriteRegisters[uiMachine - 1];
END_FOR;
FOR uiMachine := 1 TO 17 DO
	GVL_HMI.auiRobotModbusReadRegisters[uiMachine] :=
		GVL_ROBOT_MODBUS.auiReadRegisters[uiMachine - 1];
END_FOR;
GVL_HMI.xSimAxisGroupErrorAllowed := GVL_AXIS_GROUP.AxisGroup.Status.xSimErrorAllowed;
GVL_HMI.astAxisFaultStatus[1] := AXIS_X.FaultStatus;
GVL_HMI.astAxisFaultStatus[2] := AXIS_Y.FaultStatus;
GVL_HMI.astAxisFaultStatus[3] := AXIS_Z.FaultStatus;
GVL_HMI.stAxisGroupFaultStatus := GROUP_XYZ.FaultStatus;
GVL_HMI.stGripperFaultStatus := ROBOT.FaultStatus.stGripper;
GVL_HMI.stRobotFaultStatus := ROBOT.FaultStatus.stRobot;
GVL_HMI.stCellFaultStatus := CELL_MANAGER.FaultStatus;
GVL_HMI.stPointFaultStatus := ROBOT.FaultStatus.stPoint;
GVL_HMI.stMagazineFaultStatus := fbMagazine1.FaultStatus;
GVL_HMI.astMagazineFaultStatus[1] := fbMagazine1.FaultStatus;
GVL_HMI.astMagazineFaultStatus[2] := fbMagazine2.FaultStatus;
GVL_HMI.rLoadCNC_1 := GVL_STATISTIC.stStatistic.stMachineStat.rLoadCNC_1;
GVL_HMI.rLoadCNC_2 := GVL_STATISTIC.stStatistic.stMachineStat.rLoadCNC_2;
GVL_HMI.rLoadCNC_3 := GVL_STATISTIC.stStatistic.stMachineStat.rLoadCNC_3;
GVL_HMI.rRobot := GVL_STATISTIC.stStatistic.stRobotStat.rRobot;

GVL_HMI.stCellStatus := GVL_CELL_MANAGER.Status;
GVL_HMI.stCellStatus.xResetAllowed := xAlarmResetAllowed;
GVL_HMI.stCellDiag := GVL_CELL_MANAGER.Diag;
GVL_HMI.stCellError := GVL_CELL_MANAGER.Error;
GVL_HMI.stCellSafetyStatus := CELL_SAFETY.Status;
GVL_HMI.stCellSafetyDiag := CELL_SAFETY.Diag;
GVL_HMI.stCellSafetyError := CELL_SAFETY.Error;
GVL_HMI.astButtonStationIoStatus := CELL_SAFETY.astButtonStationIoStatus;
GVL_HMI.stFrontControlCabinetIoStatus := CELL_SAFETY.stFrontControlCabinetIoStatus;
GVL_HMI.xSignalTowerRed := GVL_CELL_SAFETY_IO.xSignalTowerRedOutput;
GVL_HMI.xSignalTowerAmber := GVL_CELL_SAFETY_IO.xSignalTowerAmberOutput;
GVL_HMI.xSignalTowerGreen := GVL_CELL_SAFETY_IO.xSignalTowerGreenOutput;
GVL_HMI.stRearControlCabinetIoStatus := CELL_SAFETY.stRearControlCabinetIoStatus;
GVL_HMI.stMpgIoStatus := CELL_SAFETY.stMpgIoStatus;
GVL_HMI.astEnclosureDoorStatus := CELL_SAFETY.astEnclosureDoorStatus;
GVL_HMI.stMultiType.Config := GVL_MULTI_TYPE.Config;
GVL_HMI.stMultiType.ConfigStatus := GVL_MULTI_TYPE.ConfigStatus;
GVL_HMI.stMultiType.CycleStatus := GVL_MULTI_TYPE.CycleStatus;

GVL_HMI.stRobotStatus := GVL_ROBOT.Status;
GVL_HMI.stRobotDiag := GVL_ROBOT.Diag;
GVL_HMI.stRobotError := GVL_ROBOT.Error;
GVL_HMI.stGripperDiag := GVL_ROBOT.GripperDiag;
GVL_HMI.stGripperError := GVL_ROBOT.GripperError;
GVL_HMI.stAxisGroupStatus := GVL_AXIS_GROUP.AxisGroup.Status;
GVL_HMI.stAxisGroupDiag := GVL_AXIS_GROUP.AxisGroup.Diag;
GVL_HMI.stAxisGroupError := GVL_AXIS_GROUP.AxisGroup.Error;
GVL_HMI.stMotionManagerStatus := GVL_MOTION_MANAGER.stMotionManager.Status;
GVL_HMI.stMotionManagerDiag := GVL_MOTION_MANAGER.stMotionManager.Diag;
GVL_HMI.stMotionManagerError := GVL_MOTION_MANAGER.stMotionManager.Error;
GVL_HMI.stPointManagerStatus := GVL_POINT_MANAGER.PointManager.Status;
GVL_HMI.stPointManagerDiag := GVL_POINT_MANAGER.PointManager.Diag;
GVL_HMI.stPointManagerError := GVL_POINT_MANAGER.PointManager.Error;

FOR uiMachine := 1 TO 3 DO
	GVL_HMI.astAxisStatus[uiMachine] := GVL_AXIS.arrAxis[uiMachine].Status;
	GVL_HMI.astAxisDiag[uiMachine] := GVL_AXIS.arrAxis[uiMachine].Diag;
	GVL_HMI.astAxisError[uiMachine] := GVL_AXIS.arrAxis[uiMachine].Error;
END_FOR;

GVL_HMI.stMagazineStatus := GVL_MAGAZINE.astStatus[1];
GVL_HMI.stMagazineDiag := GVL_MAGAZINE.astDiag[1];
GVL_HMI.stMagazineError := GVL_MAGAZINE.astError[1];
FOR uiMagazine := UINT#1 TO UINT#2 DO
	GVL_HMI.astMagazineStatus[uiMagazine] := GVL_MAGAZINE.astStatus[uiMagazine];
	GVL_HMI.astMagazineDiag[uiMagazine] := GVL_MAGAZINE.astDiag[uiMagazine];
	GVL_HMI.astMagazineError[uiMagazine] := GVL_MAGAZINE.astError[uiMagazine];
END_FOR;
GVL_HMI.stAlarmStatus := GVL_ALARM.Status;
IF ALARM_MANAGER.xEventsUpdated OR NOT xHmiTablesInitialized THEN
    GVL_HMI.stHmiDataRevision.udiAlarmEvents := GVL_HMI.stHmiDataRevision.udiAlarmEvents + UDINT#1;
    GVL_HMI.astAlarmEvent := GVL_ALARM.Events;
    GVL_HMI.stHmiDataRevision.udiAlarmEvents := GVL_HMI.stHmiDataRevision.udiAlarmEvents + UDINT#1;
END_IF;

FOR uiMachine := 1 TO 3 DO
	GVL_HMI.astMachineStatus[uiMachine] := GVL_MACHINE.Status[uiMachine];
	GVL_HMI.astMachineDiag[uiMachine] := GVL_MACHINE.Diag[uiMachine];
	GVL_HMI.astMachineError[uiMachine] := GVL_MACHINE.Error[uiMachine];
	CASE uiMachine OF
		1:
			GVL_HMI.astMachineFaultStatus[uiMachine] := MACHINE_1_FAULT.Status;
			GVL_HMI.astMachineFaultStatus[uiMachine].xResetAllowed :=
				MACHINE_1_SIM.Diag.xResetAllowed OR GVL_MACHINE.Status[uiMachine].xResetAllowed;
		2:
			GVL_HMI.astMachineFaultStatus[uiMachine] := MACHINE_2_FAULT.Status;
			GVL_HMI.astMachineFaultStatus[uiMachine].xResetAllowed :=
				MACHINE_2_SIM.Diag.xResetAllowed OR GVL_MACHINE.Status[uiMachine].xResetAllowed;
		3:
			GVL_HMI.astMachineFaultStatus[uiMachine] := MACHINE_3_FAULT.Status;
			GVL_HMI.astMachineFaultStatus[uiMachine].xResetAllowed :=
				MACHINE_3_SIM.Diag.xResetAllowed OR GVL_MACHINE.Status[uiMachine].xResetAllowed;
	END_CASE;
END_FOR;

GVL_HMI.astMachineIoStatus[1] := MACHINE_1_FAULT.MachineStatus;
GVL_HMI.astMachineIoStatus[2] := MACHINE_2_FAULT.MachineStatus;
GVL_HMI.astMachineIoStatus[3] := MACHINE_3_FAULT.MachineStatus;
GVL_HMI.astMachineRawIoStatus[1] := MACHINE_1_SIM.Status;
GVL_HMI.astMachineRawIoStatus[2] := MACHINE_2_SIM.Status;
GVL_HMI.astMachineRawIoStatus[3] := MACHINE_3_SIM.Status;
GVL_HMI.astMachineTimeouts[1] := MACHINE_1_FAULT.Timeouts;
GVL_HMI.astMachineTimeouts[2] := MACHINE_2_FAULT.Timeouts;
GVL_HMI.astMachineTimeouts[3] := MACHINE_3_FAULT.Timeouts;
GVL_HMI.astMachineSimDiag[1] := MACHINE_1_SIM.Diag;
GVL_HMI.astMachineSimDiag[2] := MACHINE_2_SIM.Diag;
GVL_HMI.astMachineSimDiag[3] := MACHINE_3_SIM.Diag;
GVL_HMI.astMachineSimError[1] := MACHINE_1_SIM.Error;
GVL_HMI.astMachineSimError[2] := MACHINE_2_SIM.Error;
GVL_HMI.astMachineSimError[3] := MACHINE_3_SIM.Error;

// Нечётная версия закрывает запись; gateway принимает одинаковую чётную до/после Read.
IF NOT xHmiTablesInitialized OR axMagazineInventoryChanged[1] OR axMagazineInventoryChanged[2]
OR fbMagazine1.xInventoryUpdated OR fbMagazine2.xInventoryUpdated THEN
    GVL_HMI.stHmiDataRevision.udiMagazineInventory := GVL_HMI.stHmiDataRevision.udiMagazineInventory + UDINT#1;
    GVL_HMI.astMagazineInventory := GVL_DETAIL.astMagazine;
    FOR iDetail := 1 TO GVL_CELL_SETTINGS.NumberDetail DO
        GVL_HMI.astMagazineSlot[iDetail] := GVL_DETAIL.astMagazine[1].aSlots[iDetail];
    END_FOR;
    GVL_HMI.stHmiDataRevision.udiMagazineInventory := GVL_HMI.stHmiDataRevision.udiMagazineInventory + UDINT#1;
END_IF;

// Ack only the snapshot actually dispatched through all consumers this scan.
FOR uiHmiCommandIndex := UINT#1 TO UINT#121 DO
	IF axHmiCommandConsumed[uiHmiCommandIndex] THEN
		GVL_HMI.audiHmiCommandAckSeq[uiHmiCommandIndex] := audiHmiCommandSnapshot[uiHmiCommandIndex];
	END_IF;
END_FOR;
GVL_HMI.udiCellSettingAckSeq := udiCellSettingSnapshot;

GVL_HMI.uiMagazineMode := GVL_TWO_PALLET.uiMode;
GVL_HMI.xMagazineModeAllowed := GVL_TWO_PALLET.xModeChangeAllowed;
GVL_HMI.astTwinStatus := GVL_TWO_PALLET.astStatus;
GVL_HMI.astTwinConfig := GVL_TWO_PALLET.astActiveConfig;
IF NOT xHmiTablesInitialized OR axTwinStoreChanged[1] OR axTwinStoreChanged[2] THEN
    GVL_HMI.stHmiDataRevision.udiTwinStore := GVL_HMI.stHmiDataRevision.udiTwinStore + UDINT#1;
    GVL_HMI.astTwinStore := GVL_TWO_PALLET.astStore;
    GVL_HMI.stHmiDataRevision.udiTwinStore := GVL_HMI.stHmiDataRevision.udiTwinStore + UDINT#1;
END_IF;
IF NOT xHmiTablesInitialized THEN
    GVL_HMI.stHmiDataRevision.udiEpoch := udiHmiCommandNowMs;
    IF GVL_HMI.stHmiDataRevision.udiEpoch = UDINT#0 THEN GVL_HMI.stHmiDataRevision.udiEpoch := UDINT#1; END_IF;
    GVL_HMI.stHmiDataRevision.uiVersion := UINT#1;
    xHmiTablesInitialized := TRUE;
END_IF;

(* ---- PLC_PRG.ReadHmiCommands.st ---- *)
METHOD PRIVATE ReadHmiCommands

// --- BEGIN IMPLEMENTATION ---

// Request counters belong to gateway; pulses and acknowledgements belong to PLC.
udiHmiCommandNowMs := TIME_TO_UDINT(TIME());
GVL_HMI.udiHmiCommandClockMs := udiHmiCommandNowMs;
FOR uiHmiCommandIndex := UINT#1 TO UINT#121 DO
	axHmiCommandConsumed[uiHmiCommandIndex] := FALSE;
	axHmiCommandPulse[uiHmiCommandIndex] := FALSE;
	// Mandatory low scan rearms every existing R_TRIG, including scenario events.
	IF NOT axHmiCommandWasHigh[uiHmiCommandIndex] THEN
		IF axHmiInternalPulse[uiHmiCommandIndex] THEN
			axHmiCommandPulse[uiHmiCommandIndex] := TRUE;
			axHmiInternalPulse[uiHmiCommandIndex] := FALSE;
		ELSE
			audiHmiCommandSnapshot[uiHmiCommandIndex] := GVL_HMI.audiHmiCommandSeq[uiHmiCommandIndex];
			IF (audiHmiCommandSnapshot[uiHmiCommandIndex] <> UDINT#0)
			AND (audiHmiCommandSnapshot[uiHmiCommandIndex] <> GVL_HMI.audiHmiCommandAckSeq[uiHmiCommandIndex]) THEN
				axHmiCommandConsumed[uiHmiCommandIndex] := TRUE;
				IF IsHmiCommandFresh(udiIssuedAtMs := GVL_HMI.audiHmiCommandIssuedAtMs[uiHmiCommandIndex]) THEN
					axHmiCommandPulse[uiHmiCommandIndex] := TRUE;
					GVL_HMI.auiHmiCommandResult[uiHmiCommandIndex] := UINT#1;
				ELSE
					GVL_HMI.auiHmiCommandResult[uiHmiCommandIndex] := UINT#2;
				END_IF;
			END_IF;
		END_IF;
	END_IF;
	axHmiCommandWasHigh[uiHmiCommandIndex] := axHmiCommandPulse[uiHmiCommandIndex];
END_FOR;

// Stable wire IDs; command-contract.mjs and static tests enforce this mapping.
GVL_HMI.xCellEnable := axHmiCommandPulse[1];
GVL_HMI.xCellDisable := axHmiCommandPulse[2];
GVL_HMI.xCellStart := axHmiCommandPulse[3];
GVL_HMI.xCellStop := axHmiCommandPulse[4];
GVL_HMI.xCellReset := axHmiCommandPulse[5];
GVL_HMI.xSafetyRelayReset := axHmiCommandPulse[6];
GVL_HMI.xCellOperatorCancel := axHmiCommandPulse[7];
GVL_HMI.xAlarmResetWarnings := axHmiCommandPulse[8];
GVL_HMI.xModbusSettingsApply := axHmiCommandPulse[9];
GVL_HMI.stMultiType.Command.xAutoDistribute := axHmiCommandPulse[10];
GVL_HMI.xSimAxisGroupError := axHmiCommandPulse[11];
GVL_HMI.xSimRobotWrongAction := axHmiCommandPulse[12];
GVL_HMI.xSimCellBothGrippers := axHmiCommandPulse[13];
GVL_HMI.xSimPointXOutOfLimit := axHmiCommandPulse[14];
GVL_HMI.xSimPointYOutOfLimit := axHmiCommandPulse[15];
GVL_HMI.xSimPointZOutOfLimit := axHmiCommandPulse[16];
GVL_HMI.xSimPointInvalidVelocity := axHmiCommandPulse[17];
GVL_HMI.xSimMagazineWrongOperation := axHmiCommandPulse[18];
GVL_HMI.xSimMagazineNoBlank := axHmiCommandPulse[19];
GVL_HMI.xSimMagazineNoFreeSlot := axHmiCommandPulse[20];
GVL_HMI.xSimMagazineInvalidSlot := axHmiCommandPulse[21];
GVL_HMI.xSimMagazineSlotContent := axHmiCommandPulse[22];
GVL_HMI.xSimMagazineGeometry := axHmiCommandPulse[23];
GVL_HMI.xRobotDrivesEnable := axHmiCommandPulse[24];
GVL_HMI.xRobotDrivesDisable := axHmiCommandPulse[25];
GVL_HMI.xRobotStop := axHmiCommandPulse[26];
GVL_HMI.xRobotReset := axHmiCommandPulse[27];
GVL_HMI.xTestEnvironmentApply := axHmiCommandPulse[28];
GVL_HMI.xTestSpeedProfileApply := axHmiCommandPulse[29];
GVL_HMI.xTestScenarioApply := axHmiCommandPulse[30];
GVL_HMI.xPointCheckStop := axHmiCommandPulse[31];
GVL_HMI.xRobotManualExecute := axHmiCommandPulse[32];
GVL_HMI.stMultiType.Command.xSetTypeCount := axHmiCommandPulse[33];
GVL_HMI.xCellOperatorChoice := axHmiCommandPulse[34];
GVL_HMI.stMultiType.Command.xSetMachineType := axHmiCommandPulse[35];
GVL_HMI.xRobotControlModeApply := axHmiCommandPulse[36];
GVL_HMI.stMultiType.Command.xSetSlotType := axHmiCommandPulse[37];
GVL_HMI.astAxisHmiCommand[1].xHome := axHmiCommandPulse[38];
GVL_HMI.astAxisHmiCommand[1].xMoveAbsolute := axHmiCommandPulse[39];
GVL_HMI.astAxisHmiCommand[1].xMoveRelative := axHmiCommandPulse[40];
GVL_HMI.axSimAxisJogConflict[1] := axHmiCommandPulse[41];
GVL_HMI.axMachineSimReset[1] := axHmiCommandPulse[42];
GVL_HMI.axMachineEnable[1] := axHmiCommandPulse[43];
GVL_HMI.axMachineDisable[1] := axHmiCommandPulse[44];
GVL_HMI.axMachineReset[1] := axHmiCommandPulse[45];
GVL_HMI.axMachineSetBlank[1] := axHmiCommandPulse[46];
GVL_HMI.axMachineSetDetail[1] := axHmiCommandPulse[47];
GVL_HMI.axMachineAcceptDoor[1] := axHmiCommandPulse[48];
GVL_HMI.axMachineRejectDoor[1] := axHmiCommandPulse[49];
GVL_HMI.axMachineAcceptRun[1] := axHmiCommandPulse[50];
GVL_HMI.axMachineRejectRun[1] := axHmiCommandPulse[51];
GVL_HMI.axMachineManualSafetyDoorOpen[1] := axHmiCommandPulse[52];
GVL_HMI.axMachineManualSafetyDoorClose[1] := axHmiCommandPulse[53];
GVL_HMI.axMachineManualHatchOpen[1] := axHmiCommandPulse[54];
GVL_HMI.axMachineManualHatchClose[1] := axHmiCommandPulse[55];
GVL_HMI.axMachineManualHatchUnlock[1] := axHmiCommandPulse[56];
GVL_HMI.axMachineManualHatchLock[1] := axHmiCommandPulse[57];
GVL_HMI.axMachineManualChuckOpen[1] := axHmiCommandPulse[58];
GVL_HMI.axMachineManualChuckClose[1] := axHmiCommandPulse[59];
GVL_HMI.astAxisHmiCommand[2].xHome := axHmiCommandPulse[60];
GVL_HMI.astAxisHmiCommand[2].xMoveAbsolute := axHmiCommandPulse[61];
GVL_HMI.astAxisHmiCommand[2].xMoveRelative := axHmiCommandPulse[62];
GVL_HMI.axSimAxisJogConflict[2] := axHmiCommandPulse[63];
GVL_HMI.axMachineSimReset[2] := axHmiCommandPulse[64];
GVL_HMI.axMachineEnable[2] := axHmiCommandPulse[65];
GVL_HMI.axMachineDisable[2] := axHmiCommandPulse[66];
GVL_HMI.axMachineReset[2] := axHmiCommandPulse[67];
GVL_HMI.axMachineSetBlank[2] := axHmiCommandPulse[68];
GVL_HMI.axMachineSetDetail[2] := axHmiCommandPulse[69];
GVL_HMI.axMachineAcceptDoor[2] := axHmiCommandPulse[70];
GVL_HMI.axMachineRejectDoor[2] := axHmiCommandPulse[71];
GVL_HMI.axMachineAcceptRun[2] := axHmiCommandPulse[72];
GVL_HMI.axMachineRejectRun[2] := axHmiCommandPulse[73];
GVL_HMI.axMachineManualSafetyDoorOpen[2] := axHmiCommandPulse[74];
GVL_HMI.axMachineManualSafetyDoorClose[2] := axHmiCommandPulse[75];
GVL_HMI.axMachineManualHatchOpen[2] := axHmiCommandPulse[76];
GVL_HMI.axMachineManualHatchClose[2] := axHmiCommandPulse[77];
GVL_HMI.axMachineManualHatchUnlock[2] := axHmiCommandPulse[78];
GVL_HMI.axMachineManualHatchLock[2] := axHmiCommandPulse[79];
GVL_HMI.axMachineManualChuckOpen[2] := axHmiCommandPulse[80];
GVL_HMI.axMachineManualChuckClose[2] := axHmiCommandPulse[81];
GVL_HMI.astAxisHmiCommand[3].xHome := axHmiCommandPulse[82];
GVL_HMI.astAxisHmiCommand[3].xMoveAbsolute := axHmiCommandPulse[83];
GVL_HMI.astAxisHmiCommand[3].xMoveRelative := axHmiCommandPulse[84];
GVL_HMI.axSimAxisJogConflict[3] := axHmiCommandPulse[85];
GVL_HMI.axMachineSimReset[3] := axHmiCommandPulse[86];
GVL_HMI.axMachineEnable[3] := axHmiCommandPulse[87];
GVL_HMI.axMachineDisable[3] := axHmiCommandPulse[88];
GVL_HMI.axMachineReset[3] := axHmiCommandPulse[89];
GVL_HMI.axMachineSetBlank[3] := axHmiCommandPulse[90];
GVL_HMI.axMachineSetDetail[3] := axHmiCommandPulse[91];
GVL_HMI.axMachineAcceptDoor[3] := axHmiCommandPulse[92];
GVL_HMI.axMachineRejectDoor[3] := axHmiCommandPulse[93];
GVL_HMI.axMachineAcceptRun[3] := axHmiCommandPulse[94];
GVL_HMI.axMachineRejectRun[3] := axHmiCommandPulse[95];
GVL_HMI.axMachineManualSafetyDoorOpen[3] := axHmiCommandPulse[96];
GVL_HMI.axMachineManualSafetyDoorClose[3] := axHmiCommandPulse[97];
GVL_HMI.axMachineManualHatchOpen[3] := axHmiCommandPulse[98];
GVL_HMI.axMachineManualHatchClose[3] := axHmiCommandPulse[99];
GVL_HMI.axMachineManualHatchUnlock[3] := axHmiCommandPulse[100];
GVL_HMI.axMachineManualHatchLock[3] := axHmiCommandPulse[101];
GVL_HMI.axMachineManualChuckOpen[3] := axHmiCommandPulse[102];
GVL_HMI.axMachineManualChuckClose[3] := axHmiCommandPulse[103];
GVL_HMI.astMagazineCommand[1].xEnable := axHmiCommandPulse[104];
GVL_HMI.astMagazineCommand[1].xDisable := axHmiCommandPulse[105];
GVL_HMI.astMagazineCommand[1].xStop := axHmiCommandPulse[106];
GVL_HMI.astMagazineCommand[1].xReset := axHmiCommandPulse[107];
GVL_HMI.astMagazineCommand[1].xFill := axHmiCommandPulse[108];
GVL_HMI.astMagazineCommand[1].xClear := axHmiCommandPulse[109];
GVL_HMI.astMagazineCommand[1].xApplySlot := axHmiCommandPulse[110];
GVL_HMI.astMagazineCommand[1].xApplyPitchX := axHmiCommandPulse[111];
GVL_HMI.astMagazineCommand[1].xApplyPitchY := axHmiCommandPulse[112];
GVL_HMI.astMagazineCommand[2].xEnable := axHmiCommandPulse[113];
GVL_HMI.astMagazineCommand[2].xDisable := axHmiCommandPulse[114];
GVL_HMI.astMagazineCommand[2].xStop := axHmiCommandPulse[115];
GVL_HMI.astMagazineCommand[2].xReset := axHmiCommandPulse[116];
GVL_HMI.astMagazineCommand[2].xFill := axHmiCommandPulse[117];
GVL_HMI.astMagazineCommand[2].xClear := axHmiCommandPulse[118];
GVL_HMI.astMagazineCommand[2].xApplySlot := axHmiCommandPulse[119];
GVL_HMI.astMagazineCommand[2].xApplyPitchX := axHmiCommandPulse[120];
GVL_HMI.astMagazineCommand[2].xApplyPitchY := axHmiCommandPulse[121];

(* ---- PLC_PRG.ReadHmiInputs.st ---- *)
METHOD PRIVATE ReadHmiInputs

// --- BEGIN IMPLEMENTATION ---

// HMI обязана поддерживать heartbeat. При потере связи PLC снимает только
// расширенные ручные команды; технологические проверки ниже остаются в PLC.
tonHmiWatchdog(
	IN := GVL_HMI.udiHmiHeartbeat = udiLastHmiHeartbeat,
	PT := GVL_CELL_SETTINGS.tHmiWatchdogTimeout
);
IF GVL_HMI.udiHmiHeartbeat <> udiLastHmiHeartbeat THEN
	udiLastHmiHeartbeat := GVL_HMI.udiHmiHeartbeat;
END_IF;
xHmiConnectionAlive := NOT tonHmiWatchdog.Q;

// Мобильная аренда отделена от общего HMI heartbeat. Gateway может быть жив,
// но движение обязано остановиться, если телефон перестал подтверждать аренду.
rtMobileMotionStart(CLK := GVL_HMI.xMobileMotionActive);
tonMobileMotionWatchdog(
	IN := GVL_HMI.xMobileMotionActive
		AND (GVL_HMI.udiMobileMotionHeartbeat = udiLastMobileMotionHeartbeat),
	PT := GVL_CELL_SETTINGS.tMobileMotionWatchdogTimeout
);
IF GVL_HMI.udiMobileMotionHeartbeat <> udiLastMobileMotionHeartbeat THEN
	udiLastMobileMotionHeartbeat := GVL_HMI.udiMobileMotionHeartbeat;
END_IF;
IF rtMobileMotionStart.Q THEN
	xMobileMotionLeaseActive := TRUE;
	rMobileMotionSpeedLimitPercent := LIMIT(
		REAL#0.1,
		GVL_CELL_SETTINGS.rPointCheckSpeedPercent,
		REAL#100.0
	);
END_IF;
IF xMobileMotionLeaseActive THEN
	// Во время аренды лимит разрешено только уменьшать. Повышение настройки
	// применяется уже к следующему мобильному движению.
	rMobileMotionSpeedLimitPercent := MIN(
		rMobileMotionSpeedLimitPercent,
		LIMIT(REAL#0.1, GVL_CELL_SETTINGS.rPointCheckSpeedPercent, REAL#100.0)
	);
END_IF;
xMobileMotionConnectionAlive := GVL_HMI.xMobileMotionActive
	AND NOT tonMobileMotionWatchdog.Q;
xMobileMotionStopRequest := xMobileMotionLeaseActive
	AND (NOT GVL_HMI.xMobileMotionActive
		OR NOT xMobileMotionConnectionAlive
		OR NOT xHmiConnectionAlive);
IF xMobileMotionStopRequest THEN
	// Сбрасываем вход аренды в PLC: восстановление сети не может само возобновить ход.
	GVL_HMI.xMobileMotionActive := FALSE;
	FOR uiMachine := 1 TO 3 DO
		GVL_HMI.astAxisHmiCommand[uiMachine].xJogPositive := FALSE;
		GVL_HMI.astAxisHmiCommand[uiMachine].xJogNegative := FALSE;
	END_FOR;
END_IF;
GVL_HMI.xMobileMotionLeaseAlive := xMobileMotionLeaseActive
	AND xMobileMotionConnectionAlive
	AND NOT xMobileMotionStopRequest;
GVL_HMI.rMobileMotionAppliedSpeedPercent := rMobileMotionSpeedLimitPercent;

xPointCheckRequest := FALSE;
tonPointCheckWatchdog(
	IN := GVL_HMI.udiPointCheckHeartbeat = udiLastPointCheckHeartbeat,
	PT := GVL_CELL_SETTINGS.tPointCheckWatchdogTimeout
);
IF GVL_HMI.udiPointCheckHeartbeat <> udiLastPointCheckHeartbeat THEN
	udiLastPointCheckHeartbeat := GVL_HMI.udiPointCheckHeartbeat;
END_IF;
xPointCheckConnectionAlive := (udiLastPointCheckHeartbeat <> UDINT#0) AND NOT tonPointCheckWatchdog.Q;
xPointCheckStopRequest := xPointCheckActive AND (GVL_HMI.xPointCheckStop
	OR NOT xPointCheckConnectionAlive OR NOT xHmiConnectionAlive);
// Stop is a PLC-owned one-scan event; its request counter is never cleared here.

IF GVL_HMI.rRobotManualSpeedPercent < REAL#0.1 THEN
	GVL_HMI.rRobotManualSpeedPercent := REAL#0.1;
ELSIF GVL_HMI.rRobotManualSpeedPercent > REAL#100.0 THEN
	GVL_HMI.rRobotManualSpeedPercent := REAL#100.0;
END_IF;
IF (GVL_HMI.lrRobotManualStep <> 0.1)
AND (GVL_HMI.lrRobotManualStep <> 1.0)
AND (GVL_HMI.lrRobotManualStep <> 10.0)
AND (GVL_HMI.lrRobotManualStep <> 100.0) THEN
	GVL_HMI.lrRobotManualStep := 1.0;
END_IF;

IF NOT xHmiConnectionAlive THEN
	FOR uiMachine := 1 TO 3 DO
		GVL_HMI.astAxisHmiCommand[uiMachine].xJogPositive := FALSE;
		GVL_HMI.astAxisHmiCommand[uiMachine].xJogNegative := FALSE;
		GVL_HMI.astAxisHmiCommand[uiMachine].xHome := FALSE;
		GVL_HMI.astAxisHmiCommand[uiMachine].xMoveAbsolute := FALSE;
		GVL_HMI.astAxisHmiCommand[uiMachine].xMoveRelative := FALSE;
	END_FOR;
	FOR uiMagazine := UINT#1 TO UINT#2 DO
		GVL_HMI.astMagazineCommand[uiMagazine].xStop := FALSE;
	END_FOR;
	GVL_HMI.xRobotManualExecute := FALSE;
END_IF;

// Глобальные команды ячейки поступают через единый интерфейс HMI.
GVL_CELL_CONTROL.xEnable := GVL_HMI.xCellEnable;
GVL_CELL_CONTROL.xDisable := GVL_HMI.xCellDisable;
GVL_CELL_CONTROL.xStart := GVL_HMI.xCellStart;
GVL_CELL_CONTROL.xStop := GVL_HMI.xCellStop;
// Необработанный общий импульс передаётся всем владельцам аварий.
// Каждый функциональный блок самостоятельно проверяет возможность сброса.
GVL_CELL_CONTROL.xReset := GVL_HMI.xCellReset;
// Режим хранит PLC. Новая транзакция применяется в RunSafety после чтения
// актуальных входов безопасности; PublishHmi не пишет в буфер запроса.
GVL_ALARM.Command.xResetWarnings := GVL_HMI.xAlarmResetWarnings;

// Режим инъекции ошибок включается отдельным переключателем страницы CELL_SETTINGS.
GVL_CELL_SETTINGS.xErrorSimulationEnabled := GVL_HMI.xErrorSimulationEnable
	AND (GVL_CELL_SETTINGS.eTestEnvironment <> E_CELL_TEST_ENVIRONMENT.NORMAL);

// Ползунок меняет только запрошенное значение. Отдельный FB применяет его к
// таймерам и Dynamic Limits безопасной транзакцией перед следующим тестом.
GVL_CELL_SETTINGS.xSimulationAccelerationChangeAllowed :=
	xHmiConnectionAlive
	AND NOT GVL_CELL_CONTROL.xGlobalError;

IF GVL_CELL_SETTINGS.xSimulationAccelerationChangeAllowed THEN
	GVL_CELL_SETTINGS.xSimulationAccelerationEnable := GVL_HMI.xSimulationAccelerationEnable;
	GVL_CELL_SETTINGS.uiSimulationTimeFactor := GVL_HMI.uiSimulationTimeFactor;
	IF GVL_CELL_SETTINGS.uiSimulationTimeFactor < UINT#1 THEN
		GVL_CELL_SETTINGS.uiSimulationTimeFactor := UINT#1;
	ELSIF GVL_CELL_SETTINGS.uiSimulationTimeFactor > UINT#100 THEN
		GVL_CELL_SETTINGS.uiSimulationTimeFactor := UINT#100;
	END_IF;
ELSE
	// При потере разрешения сохраняем последнее принятое требование.
	GVL_HMI.xSimulationAccelerationEnable := GVL_CELL_SETTINGS.xSimulationAccelerationActive;
	GVL_HMI.uiSimulationTimeFactor := GVL_CELL_SETTINGS.uiSimulationTimeFactor;
END_IF;

// Общие технологические TIMEOUT и допуски HOME принимаются только при полностью
// остановленной ячейке. Координатами HOME_SAFETY владеет редактор точек ниже.
GVL_CELL_SETTINGS.xCellSettingsChangeAllowed :=
	xHmiConnectionAlive
	AND NOT GVL_CELL_MANAGER.Status.xRunning
	AND NOT GVL_HMI.xModbusMode
	AND NOT GVL_CELL_CONTROL.xGlobalError
	AND NOT GVL_AXIS.arrAxis[1].Status.xMotionBusy
	AND NOT GVL_AXIS.arrAxis[2].Status.xMotionBusy
	AND NOT GVL_AXIS.arrAxis[3].Status.xMotionBusy
	AND NOT GVL_AXIS_GROUP.AxisGroup.Command.xMoveDirect
	AND NOT GVL_AXIS_GROUP.AxisGroup.Command.xMoveLinear
	AND NOT xPowerTransitionActive
	AND NOT SIMULATION_DYNAMICS.xBusy
	AND NOT GVL_ROBOT.Status.xBusy;

GVL_CELL_SETTINGS.xIoFilterSettingsChangeAllowed := xHmiConnectionAlive
	AND GVL_CELL_CONTROL.xManual
	AND NOT GVL_CELL_MANAGER.Status.xRunning
	AND NOT GVL_ROBOT.Status.xBusy AND NOT xMotionBusy
	AND NOT xPowerTransitionActive AND NOT SIMULATION_DYNAMICS.xBusy
	AND NOT GVL_MACHINE.Status[1].xBusy AND NOT GVL_MACHINE.Status[1].xProcessing
	AND NOT GVL_MACHINE.Status[2].xBusy AND NOT GVL_MACHINE.Status[2].xProcessing
	AND NOT GVL_MACHINE.Status[3].xBusy AND NOT GVL_MACHINE.Status[3].xProcessing
	AND NOT GVL_TWO_PALLET.astStatus[1].xBusy AND NOT GVL_TWO_PALLET.astStatus[2].xBusy
	AND NOT GVL_TWO_PALLET.astInput[1].xPowered AND NOT GVL_TWO_PALLET.astInput[2].xPowered;

// Допуск принадлежит конкретному магазину; общий редактор не обходит занятость зоны.
FOR uiCalibrationMagazine := UINT#1 TO UINT#2 DO
	xMagazineCalibrationEditAllowed[uiCalibrationMagazine] :=
		NOT GVL_MAGAZINE.astStatus[uiCalibrationMagazine].xEnabled
		AND NOT GVL_MAGAZINE.astStatus[uiCalibrationMagazine].xBusy
		AND NOT GVL_TWO_PALLET.astStatus[uiCalibrationMagazine].xEnabled
		AND NOT GVL_TWO_PALLET.astStatus[uiCalibrationMagazine].xBusy
		AND (GVL_ROBOT.Status.uiMagazineContext <> uiCalibrationMagazine);
	GVL_HMI.astMagazineCalibrationStatus[uiCalibrationMagazine].xChangeAllowed :=
		GVL_CELL_SETTINGS.xCellSettingsChangeAllowed
		AND xMagazineCalibrationEditAllowed[uiCalibrationMagazine]
		AND NOT xPointCheckActive;
END_FOR;

// Independent requested value; publication cannot overwrite an incoming write.
xCellSettingRejected := FALSE;
udiCellSettingSnapshot := GVL_HMI.udiCellSettingCommandSeq;
IF (udiCellSettingSnapshot <> UDINT#0)
AND (udiCellSettingSnapshot <> GVL_HMI.udiCellSettingAckSeq) THEN
	GVL_HMI.uiCellSettingResult := UINT#3;
	IF NOT IsHmiCommandFresh(udiIssuedAtMs := GVL_HMI.udiCellSettingIssuedAtMs) THEN
		GVL_HMI.uiCellSettingResult := UINT#4; // Expired: never apply later
	ELSIF ((((GVL_HMI.uiCellSettingIndex = UINT#37) OR (GVL_HMI.uiCellSettingIndex = UINT#38) OR (GVL_HMI.uiCellSettingIndex = UINT#39))
		AND NOT GVL_CELL_SETTINGS.xIoFilterSettingsChangeAllowed)
		OR (((GVL_HMI.uiCellSettingIndex <> UINT#37) AND (GVL_HMI.uiCellSettingIndex <> UINT#38) AND (GVL_HMI.uiCellSettingIndex <> UINT#39))
			AND NOT GVL_CELL_SETTINGS.xCellSettingsChangeAllowed))
	OR (((GVL_HMI.uiCellSettingIndex = UINT#4)
		OR (GVL_HMI.uiCellSettingIndex = UINT#25)
		OR (GVL_HMI.uiCellSettingIndex = UINT#29))
		AND xPointCheckActive)
	OR ((GVL_HMI.uiCellSettingIndex = UINT#28) AND xMobileMotionLeaseActive) THEN
		GVL_HMI.uiCellSettingResult := UINT#2;
	ELSE
		CASE GVL_HMI.uiCellSettingIndex OF
			UINT#1:
				IF (GVL_HMI.lrCellSettingRequest >= 0.1) AND (GVL_HMI.lrCellSettingRequest <= 1000.0) THEN
					GVL_CELL_SETTINGS.lrSafetyHomeToleranceX := GVL_HMI.lrCellSettingRequest;
					GVL_HMI.uiCellSettingResult := UINT#1;
				END_IF;
			UINT#2:
				IF (GVL_HMI.lrCellSettingRequest >= 0.1) AND (GVL_HMI.lrCellSettingRequest <= 1000.0) THEN
					GVL_CELL_SETTINGS.lrSafetyHomeToleranceY := GVL_HMI.lrCellSettingRequest;
					GVL_HMI.uiCellSettingResult := UINT#1;
				END_IF;
			UINT#3:
				IF (GVL_HMI.lrCellSettingRequest >= 0.1) AND (GVL_HMI.lrCellSettingRequest <= 1000.0) THEN
					GVL_CELL_SETTINGS.lrSafetyHomeToleranceZ := GVL_HMI.lrCellSettingRequest;
					GVL_HMI.uiCellSettingResult := UINT#1;
				END_IF;
			UINT#4:
				IF (GVL_HMI.lrCellSettingRequest >= 0.1) AND (GVL_HMI.lrCellSettingRequest <= 100.0) THEN
					GVL_CELL_SETTINGS.rPointCheckSpeedPercent := LREAL_TO_REAL(GVL_HMI.lrCellSettingRequest);
					GVL_HMI.uiCellSettingResult := UINT#1;
				END_IF;
			UINT#5:
				IF (GVL_HMI.lrCellSettingRequest >= 1000.0) AND (GVL_HMI.lrCellSettingRequest <= 600000.0) THEN
					GVL_CELL_SETTINGS.stMachineTimeouts.tRobotMove := UDINT_TO_TIME(LREAL_TO_UDINT(GVL_HMI.lrCellSettingRequest));
					GVL_HMI.uiCellSettingResult := UINT#1;
				END_IF;
			UINT#6:
				IF (GVL_HMI.lrCellSettingRequest >= 1000.0) AND (GVL_HMI.lrCellSettingRequest <= 600000.0) THEN
					GVL_CELL_SETTINGS.stMachineTimeouts.tRobotAction := UDINT_TO_TIME(LREAL_TO_UDINT(GVL_HMI.lrCellSettingRequest));
					GVL_HMI.uiCellSettingResult := UINT#1;
				END_IF;
			UINT#7:
				IF (GVL_HMI.lrCellSettingRequest >= 1000.0) AND (GVL_HMI.lrCellSettingRequest <= 600000.0) THEN
					GVL_CELL_SETTINGS.stMachineTimeouts.tRobotRelease := UDINT_TO_TIME(LREAL_TO_UDINT(GVL_HMI.lrCellSettingRequest));
					GVL_HMI.uiCellSettingResult := UINT#1;
				END_IF;
			UINT#8:
				IF (GVL_HMI.lrCellSettingRequest >= 1000.0) AND (GVL_HMI.lrCellSettingRequest <= 600000.0) THEN
					GVL_CELL_SETTINGS.stMachineTimeouts.tDoorOpen := UDINT_TO_TIME(LREAL_TO_UDINT(GVL_HMI.lrCellSettingRequest));
					GVL_HMI.uiCellSettingResult := UINT#1;
				END_IF;
			UINT#9:
				IF (GVL_HMI.lrCellSettingRequest >= 1000.0) AND (GVL_HMI.lrCellSettingRequest <= 600000.0) THEN
					GVL_CELL_SETTINGS.stMachineTimeouts.tDoorClose := UDINT_TO_TIME(LREAL_TO_UDINT(GVL_HMI.lrCellSettingRequest));
					GVL_HMI.uiCellSettingResult := UINT#1;
				END_IF;
			UINT#10:
				IF (GVL_HMI.lrCellSettingRequest >= 1000.0) AND (GVL_HMI.lrCellSettingRequest <= 600000.0) THEN
					GVL_CELL_SETTINGS.stMachineTimeouts.tHatchUnlock := UDINT_TO_TIME(LREAL_TO_UDINT(GVL_HMI.lrCellSettingRequest));
					GVL_HMI.uiCellSettingResult := UINT#1;
				END_IF;
			UINT#11:
				IF (GVL_HMI.lrCellSettingRequest >= 1000.0) AND (GVL_HMI.lrCellSettingRequest <= 600000.0) THEN
					GVL_CELL_SETTINGS.stMachineTimeouts.tChuckOpen := UDINT_TO_TIME(LREAL_TO_UDINT(GVL_HMI.lrCellSettingRequest));
					GVL_HMI.uiCellSettingResult := UINT#1;
				END_IF;
			UINT#12:
				IF (GVL_HMI.lrCellSettingRequest >= 1000.0) AND (GVL_HMI.lrCellSettingRequest <= 600000.0) THEN
					GVL_CELL_SETTINGS.stMachineTimeouts.tChuckClose := UDINT_TO_TIME(LREAL_TO_UDINT(GVL_HMI.lrCellSettingRequest));
					GVL_HMI.uiCellSettingResult := UINT#1;
				END_IF;
			UINT#13:
				IF (GVL_HMI.lrCellSettingRequest >= 1000.0) AND (GVL_HMI.lrCellSettingRequest <= 600000.0) THEN
					GVL_CELL_SETTINGS.stMachineTimeouts.tCycleStart := UDINT_TO_TIME(LREAL_TO_UDINT(GVL_HMI.lrCellSettingRequest));
					GVL_HMI.uiCellSettingResult := UINT#1;
				END_IF;
			UINT#14:
				IF (GVL_HMI.lrCellSettingRequest >= 1000.0) AND (GVL_HMI.lrCellSettingRequest <= 600000.0) THEN
					GVL_CELL_SETTINGS.stAxisTimeouts.tPowerTimeout := UDINT_TO_TIME(LREAL_TO_UDINT(GVL_HMI.lrCellSettingRequest));
					GVL_HMI.uiCellSettingResult := UINT#1;
				END_IF;
			UINT#15:
				IF (GVL_HMI.lrCellSettingRequest >= 1000.0) AND (GVL_HMI.lrCellSettingRequest <= 600000.0) THEN
					GVL_CELL_SETTINGS.stAxisTimeouts.tResetTimeout := UDINT_TO_TIME(LREAL_TO_UDINT(GVL_HMI.lrCellSettingRequest));
					GVL_HMI.uiCellSettingResult := UINT#1;
				END_IF;
			UINT#16:
				IF (GVL_HMI.lrCellSettingRequest >= 1000.0) AND (GVL_HMI.lrCellSettingRequest <= 600000.0) THEN
					GVL_CELL_SETTINGS.stAxisTimeouts.tStopTimeout := UDINT_TO_TIME(LREAL_TO_UDINT(GVL_HMI.lrCellSettingRequest));
					GVL_HMI.uiCellSettingResult := UINT#1;
				END_IF;
			UINT#17:
				IF (GVL_HMI.lrCellSettingRequest >= 1000.0) AND (GVL_HMI.lrCellSettingRequest <= 600000.0) THEN
					GVL_CELL_SETTINGS.stAxisTimeouts.tHomeTimeout := UDINT_TO_TIME(LREAL_TO_UDINT(GVL_HMI.lrCellSettingRequest));
					GVL_HMI.uiCellSettingResult := UINT#1;
				END_IF;
			UINT#18:
				IF (GVL_HMI.lrCellSettingRequest >= 1000.0) AND (GVL_HMI.lrCellSettingRequest <= 600000.0) THEN
					GVL_CELL_SETTINGS.stAxisTimeouts.tMoveTimeout := UDINT_TO_TIME(LREAL_TO_UDINT(GVL_HMI.lrCellSettingRequest));
					GVL_HMI.uiCellSettingResult := UINT#1;
				END_IF;
			UINT#19:
				IF (GVL_HMI.lrCellSettingRequest >= 1000.0) AND (GVL_HMI.lrCellSettingRequest <= 600000.0) THEN
					GVL_CELL_SETTINGS.stAxisGroupTimeouts.tPowerTimeout := UDINT_TO_TIME(LREAL_TO_UDINT(GVL_HMI.lrCellSettingRequest));
					GVL_HMI.uiCellSettingResult := UINT#1;
				END_IF;
			UINT#20:
				IF (GVL_HMI.lrCellSettingRequest >= 1000.0) AND (GVL_HMI.lrCellSettingRequest <= 600000.0) THEN
					GVL_CELL_SETTINGS.stAxisGroupTimeouts.tGroupTimeout := UDINT_TO_TIME(LREAL_TO_UDINT(GVL_HMI.lrCellSettingRequest));
					GVL_HMI.uiCellSettingResult := UINT#1;
				END_IF;
			UINT#21:
				IF (GVL_HMI.lrCellSettingRequest >= 1000.0) AND (GVL_HMI.lrCellSettingRequest <= 600000.0) THEN
					GVL_CELL_SETTINGS.stAxisGroupTimeouts.tStopTimeout := UDINT_TO_TIME(LREAL_TO_UDINT(GVL_HMI.lrCellSettingRequest));
					GVL_HMI.uiCellSettingResult := UINT#1;
				END_IF;
			UINT#22:
				IF (GVL_HMI.lrCellSettingRequest >= 1000.0) AND (GVL_HMI.lrCellSettingRequest <= 600000.0) THEN
					GVL_CELL_SETTINGS.stAxisGroupTimeouts.tHaltTimeout := UDINT_TO_TIME(LREAL_TO_UDINT(GVL_HMI.lrCellSettingRequest));
					GVL_HMI.uiCellSettingResult := UINT#1;
				END_IF;
			UINT#23:
				IF (GVL_HMI.lrCellSettingRequest >= 1000.0) AND (GVL_HMI.lrCellSettingRequest <= 600000.0) THEN
					GVL_CELL_SETTINGS.stAxisGroupTimeouts.tHomeTimeout := UDINT_TO_TIME(LREAL_TO_UDINT(GVL_HMI.lrCellSettingRequest));
					GVL_HMI.uiCellSettingResult := UINT#1;
				END_IF;
			UINT#24:
				IF (GVL_HMI.lrCellSettingRequest >= 1000.0) AND (GVL_HMI.lrCellSettingRequest <= 600000.0) THEN
					GVL_CELL_SETTINGS.stAxisGroupTimeouts.tMoveTimeout := UDINT_TO_TIME(LREAL_TO_UDINT(GVL_HMI.lrCellSettingRequest));
					GVL_HMI.uiCellSettingResult := UINT#1;
				END_IF;
			UINT#25:
				IF (GVL_HMI.lrCellSettingRequest >= 500.0) AND (GVL_HMI.lrCellSettingRequest <= 60000.0) THEN
					GVL_CELL_SETTINGS.tPointCheckStartTimeout := UDINT_TO_TIME(LREAL_TO_UDINT(GVL_HMI.lrCellSettingRequest));
					GVL_HMI.uiCellSettingResult := UINT#1;
				END_IF;
			UINT#26:
				IF (GVL_HMI.lrCellSettingRequest >= 1000.0) AND (GVL_HMI.lrCellSettingRequest <= 600000.0) THEN
					GVL_CELL_SETTINGS.tSimulationDynamicsTimeout := UDINT_TO_TIME(LREAL_TO_UDINT(GVL_HMI.lrCellSettingRequest));
					GVL_HMI.uiCellSettingResult := UINT#1;
				END_IF;
			UINT#27:
				IF (GVL_HMI.lrCellSettingRequest >= 500.0) AND (GVL_HMI.lrCellSettingRequest <= 30000.0) THEN
					GVL_CELL_SETTINGS.tHmiWatchdogTimeout := UDINT_TO_TIME(LREAL_TO_UDINT(GVL_HMI.lrCellSettingRequest));
					GVL_HMI.uiCellSettingResult := UINT#1;
				END_IF;
			UINT#28:
				IF (GVL_HMI.lrCellSettingRequest >= 500.0) AND (GVL_HMI.lrCellSettingRequest <= 30000.0) THEN
					GVL_CELL_SETTINGS.tMobileMotionWatchdogTimeout := UDINT_TO_TIME(LREAL_TO_UDINT(GVL_HMI.lrCellSettingRequest));
					GVL_HMI.uiCellSettingResult := UINT#1;
				END_IF;
			UINT#29:
				IF (GVL_HMI.lrCellSettingRequest >= 500.0) AND (GVL_HMI.lrCellSettingRequest <= 30000.0) THEN
					GVL_CELL_SETTINGS.tPointCheckWatchdogTimeout := UDINT_TO_TIME(LREAL_TO_UDINT(GVL_HMI.lrCellSettingRequest));
					GVL_HMI.uiCellSettingResult := UINT#1;
				END_IF;
			UINT#30:
				IF (GVL_HMI.lrCellSettingRequest >= 1000.0) AND (GVL_HMI.lrCellSettingRequest <= 30000.0) THEN
					GVL_CELL_SETTINGS.tHmiCommandFreshnessTimeout := UDINT_TO_TIME(LREAL_TO_UDINT(GVL_HMI.lrCellSettingRequest));
					GVL_HMI.uiCellSettingResult := UINT#1;
				END_IF;
			UINT#31:
				IF (GVL_HMI.lrCellSettingRequest >= 100.0) AND (GVL_HMI.lrCellSettingRequest <= 10000.0) THEN
					GVL_CELL_SETTINGS.stAxisTimeouts.tPowerFeedbackLossTimeout := UDINT_TO_TIME(LREAL_TO_UDINT(GVL_HMI.lrCellSettingRequest));
					GVL_HMI.uiCellSettingResult := UINT#1;
				END_IF;
			UINT#32:
				IF (GVL_HMI.lrCellSettingRequest >= 1.0) AND (GVL_HMI.lrCellSettingRequest <= 100.0) THEN
					GVL_CELL_SETTINGS.rRobotAccelerationPercent := LREAL_TO_REAL(GVL_HMI.lrCellSettingRequest);
					GVL_HMI.uiCellSettingResult := UINT#1;
				END_IF;
			UINT#33:
				IF (GVL_HMI.lrCellSettingRequest >= 1.0) AND (GVL_HMI.lrCellSettingRequest <= 100.0) THEN
					GVL_CELL_SETTINGS.rRobotDecelerationPercent := LREAL_TO_REAL(GVL_HMI.lrCellSettingRequest);
					GVL_HMI.uiCellSettingResult := UINT#1;
				END_IF;
			UINT#34:
				IF (GVL_HMI.lrCellSettingRequest >= 1.0) AND (GVL_HMI.lrCellSettingRequest <= 100.0) THEN
					GVL_CELL_SETTINGS.rRobotJerkPercent := LREAL_TO_REAL(GVL_HMI.lrCellSettingRequest);
					GVL_HMI.uiCellSettingResult := UINT#1;
				END_IF;
			UINT#35:
				IF (GVL_HMI.lrCellSettingRequest >= 1.0) AND (GVL_HMI.lrCellSettingRequest <= 100000.0) THEN
					GVL_CELL_SETTINGS.lrRobotHaltDeceleration := GVL_HMI.lrCellSettingRequest;
					GVL_HMI.uiCellSettingResult := UINT#1;
				END_IF;
			UINT#36:
				IF (GVL_HMI.lrCellSettingRequest >= 1.0) AND (GVL_HMI.lrCellSettingRequest <= 1000000.0) THEN
					GVL_CELL_SETTINGS.lrRobotHaltJerk := GVL_HMI.lrCellSettingRequest;
					GVL_HMI.uiCellSettingResult := UINT#1;
				END_IF;
			UINT#37:
				IF (GVL_HMI.lrCellSettingRequest >= 0.0) AND (GVL_HMI.lrCellSettingRequest <= 5000.0) THEN
					GVL_CELL_SETTINGS.tInputFilterRise := UDINT_TO_TIME(LREAL_TO_UDINT(GVL_HMI.lrCellSettingRequest));
					GVL_HMI.uiCellSettingResult := UINT#1;
				END_IF;
			UINT#38:
				IF (GVL_HMI.lrCellSettingRequest >= 0.0) AND (GVL_HMI.lrCellSettingRequest <= 5000.0) THEN
					GVL_CELL_SETTINGS.tInputFilterFall := UDINT_TO_TIME(LREAL_TO_UDINT(GVL_HMI.lrCellSettingRequest));
					GVL_HMI.uiCellSettingResult := UINT#1;
				END_IF;
			UINT#39:
				IF (GVL_HMI.lrCellSettingRequest >= 0.0) AND (GVL_HMI.lrCellSettingRequest <= 60000.0) THEN
					GVL_CELL_SETTINGS.tAlarmHornDuration := UDINT_TO_TIME(LREAL_TO_UDINT(GVL_HMI.lrCellSettingRequest));
					GVL_HMI.uiCellSettingResult := UINT#1;
				END_IF;
			UINT#40, UINT#41:
				uiCalibrationSettingMagazine := GVL_HMI.uiCellSettingIndex - UINT#39;
				IF NOT GVL_HMI.astMagazineCalibrationStatus[uiCalibrationSettingMagazine].xChangeAllowed THEN
					GVL_HMI.uiCellSettingResult := UINT#2;
				ELSIF (GVL_HMI.lrCellSettingRequest = 1.0) OR (GVL_HMI.lrCellSettingRequest = 3.0) THEN
					IF Persistent_Value.astMagazineCalibration[uiCalibrationSettingMagazine].uiMethod <> LREAL_TO_UINT(GVL_HMI.lrCellSettingRequest) THEN
						Persistent_Value.astMagazineCalibration[uiCalibrationSettingMagazine].uiMethod := LREAL_TO_UINT(GVL_HMI.lrCellSettingRequest);
						InvalidateMagazineCalibration(uiMagazine := uiCalibrationSettingMagazine);
					END_IF;
					GVL_HMI.uiCellSettingResult := UINT#1;
				END_IF;
		END_CASE;
	END_IF;
	xCellSettingRejected := GVL_HMI.uiCellSettingResult <> UINT#1;
END_IF;

// =============================================================================
// Транзакционный редактор 18 фиксированных инженерных точек
// =============================================================================
xPointEditorAllHomed := GVL_AXIS.arrAxis[1].Status.xHomed
	AND GVL_AXIS.arrAxis[2].Status.xHomed
	AND GVL_AXIS.arrAxis[3].Status.xHomed;
xPointEditorBaseAllowed := xHmiConnectionAlive
	AND NOT xPointCheckActive
	AND GVL_CELL_CONTROL.xManual
	AND NOT GVL_HMI.xModbusMode
	AND NOT GVL_CELL_MANAGER.Status.xRunning
	AND NOT GVL_CELL_CONTROL.xGlobalError
	AND NOT GVL_ROBOT.Status.xBusy
	AND NOT xMotionBusy
	AND NOT xDriveError
	AND NOT GVL_MOTION_MANAGER.stMotionManager.Status.xError
	AND xPointEditorAllHomed
	AND GVL_AXIS_GROUP.AxisGroup.Status.xPositionValid;
GVL_HMI.xPointEditorCaptureAllowed := xPointEditorBaseAllowed;
GVL_HMI.xPointEditorSaveAllowed := xPointEditorBaseAllowed
	AND GVL_POINT_MANAGER.PointManager.Diag.xXLimitValid
	AND GVL_POINT_MANAGER.PointManager.Diag.xYLimitValid
	AND GVL_POINT_MANAGER.PointManager.Diag.xZLimitValid;
FOR uiCalibrationMagazine := UINT#1 TO UINT#2 DO
	GVL_HMI.astMagazineCalibrationStatus[uiCalibrationMagazine].xCaptureAllowed :=
		GVL_HMI.xPointEditorCaptureAllowed;
	GVL_HMI.astMagazineCalibrationStatus[uiCalibrationMagazine].xSaveAllowed :=
		GVL_HMI.xPointEditorSaveAllowed;
	GVL_HMI.astMagazineCalibrationStatus[uiCalibrationMagazine].xReferenceCaptureAllowed :=
		GVL_HMI.astMagazineCalibrationStatus[uiCalibrationMagazine].xCaptureAllowed
		AND (Persistent_Value.astMagazineCalibration[uiCalibrationMagazine].uiMethod = UINT#3);
	GVL_HMI.astMagazineCalibrationStatus[uiCalibrationMagazine].xReferenceSaveAllowed :=
		GVL_HMI.astMagazineCalibrationStatus[uiCalibrationMagazine].xSaveAllowed
		AND (Persistent_Value.astMagazineCalibration[uiCalibrationMagazine].uiMethod = UINT#3);
END_FOR;

IF (GVL_HMI.udiPointEditorCommandSeq <> UDINT#0)
AND (GVL_HMI.udiPointEditorCommandSeq <> udiLastPointEditorCommandSeq) THEN
	udiLastPointEditorCommandSeq := GVL_HMI.udiPointEditorCommandSeq;
	GVL_HMI.uiPointEditorResult := UINT#2;
	GVL_HMI.uiPointEditorRejectReason := UINT#0;
	xPointEditorRequestValid := FALSE;
	xPointEditorMagazinePoint := FALSE;
	uiPointEditorGeometryStation := UINT#0;
	uiPointEditorMagazine := UINT#0;
	uiPointEditorReference := UINT#0;
	ePointEditorName := E_POINT_NAME.NONE;
	uiPointStorageIndex := UINT#0;

	CASE GVL_HMI.uiPointEditorIndex OF
		UINT#1: ePointEditorName := E_POINT_NAME.MACHINE_1_ABOVE; uiPointStorageIndex := UINT#1;
		UINT#2: ePointEditorName := E_POINT_NAME.MACHINE_1_CHUCK_APROACH; uiPointStorageIndex := UINT#3;
		UINT#3: ePointEditorName := E_POINT_NAME.MACHINE_1_CHUCK_POSITION; uiPointStorageIndex := UINT#4;
		UINT#4: ePointEditorName := E_POINT_NAME.MACHINE_2_ABOVE; uiPointStorageIndex := UINT#5;
		UINT#5: ePointEditorName := E_POINT_NAME.MACHINE_2_CHUCK_APROACH; uiPointStorageIndex := UINT#7;
		UINT#6: ePointEditorName := E_POINT_NAME.MACHINE_2_CHUCK_POSITION; uiPointStorageIndex := UINT#8;
		UINT#7: ePointEditorName := E_POINT_NAME.MACHINE_3_ABOVE; uiPointStorageIndex := UINT#9;
		UINT#8: ePointEditorName := E_POINT_NAME.MACHINE_3_CHUCK_APROACH; uiPointStorageIndex := UINT#11;
		UINT#9: ePointEditorName := E_POINT_NAME.MACHINE_3_CHUCK_POSITION; uiPointStorageIndex := UINT#12;
		UINT#10: ePointEditorName := E_POINT_NAME.HOME_SAFETY; uiPointStorageIndex := UINT#13;
		UINT#11: ePointEditorName := E_POINT_NAME.MAGAZINE_1_DETAIL; uiPointStorageIndex := UINT#14; uiPointEditorMagazine := UINT#1;
		UINT#12: ePointEditorName := E_POINT_NAME.MAGAZINE_2_DETAIL; uiPointStorageIndex := UINT#15; uiPointEditorMagazine := UINT#2;
		UINT#13: ePointEditorName := E_POINT_NAME.GEOMETRY_1_PLACE; uiPointEditorGeometryStation := UINT#1;
		UINT#14: ePointEditorName := E_POINT_NAME.GEOMETRY_2_PLACE; uiPointEditorGeometryStation := UINT#2;
		UINT#15: ePointEditorName := E_POINT_NAME.MAGAZINE_1_AXIS_X; uiPointEditorMagazine := UINT#1; uiPointEditorReference := UINT#1;
		UINT#16: ePointEditorName := E_POINT_NAME.MAGAZINE_1_AXIS_Y; uiPointEditorMagazine := UINT#1; uiPointEditorReference := UINT#2;
		UINT#17: ePointEditorName := E_POINT_NAME.MAGAZINE_2_AXIS_X; uiPointEditorMagazine := UINT#2; uiPointEditorReference := UINT#1;
		UINT#18: ePointEditorName := E_POINT_NAME.MAGAZINE_2_AXIS_Y; uiPointEditorMagazine := UINT#2; uiPointEditorReference := UINT#2;
	END_CASE;
	xPointEditorRequestValid := (ePointEditorName <> E_POINT_NAME.NONE)
		AND ((uiPointStorageIndex <> UINT#0) OR (uiPointEditorGeometryStation <> UINT#0)
			OR (uiPointEditorReference <> UINT#0));
	xPointEditorMagazinePoint := (ePointEditorName = E_POINT_NAME.MAGAZINE_1_DETAIL)
		OR (ePointEditorName = E_POINT_NAME.MAGAZINE_2_DETAIL);
	xPointEditorGeometrySave := (GVL_HMI.uiPointEditorCommand = UINT#2)
		AND (uiPointEditorGeometryStation <> UINT#0);

	IF (GVL_HMI.uiPointEditorCommand <> UINT#1)
	AND (GVL_HMI.uiPointEditorCommand <> UINT#2)
	AND (GVL_HMI.uiPointEditorCommand <> UINT#3)
	AND (GVL_HMI.uiPointEditorCommand <> UINT#4) THEN
		GVL_HMI.uiPointEditorRejectReason := UINT#1; // Неизвестная команда
	ELSIF NOT xPointEditorRequestValid
	OR ((GVL_HMI.uiPointEditorCommand = UINT#4) AND NOT xPointEditorMagazinePoint) THEN
		GVL_HMI.uiPointEditorRejectReason := UINT#2; // Неверный индекс точки
	ELSIF NOT xHmiConnectionAlive THEN
		GVL_HMI.uiPointEditorRejectReason := UINT#3; // HMI offline
	ELSIF xPointEditorGeometrySave THEN
		// SAVE только изменяет данные. Режим, Home, движение, ошибки и состояние
		// ГК не блокируют запись. CAPTURE/CHECK сохраняют прежние допуски.
		IF GVL_HMI.xModbusMode
		OR (GVL_CELL_SETTINGS.eTestEnvironment = E_CELL_TEST_ENVIRONMENT.SC500_BENCH) THEN
			GVL_HMI.uiPointEditorRejectReason := UINT#5;
		ELSIF NOT GVL_POINT_MANAGER.PointManager.Diag.xXLimitValid
		OR NOT GVL_POINT_MANAGER.PointManager.Diag.xYLimitValid
		OR NOT GVL_POINT_MANAGER.PointManager.Diag.xZLimitValid THEN
			GVL_HMI.uiPointEditorRejectReason := UINT#13;
		END_IF;
	ELSIF NOT GVL_CELL_CONTROL.xManual THEN
		GVL_HMI.uiPointEditorRejectReason := UINT#4; // Требуется ручной режим
	ELSIF GVL_HMI.xModbusMode THEN
		GVL_HMI.uiPointEditorRejectReason := UINT#5; // Требуется SoftMotion
	ELSIF GVL_CELL_MANAGER.Status.xRunning THEN
		GVL_HMI.uiPointEditorRejectReason := UINT#6; // Автоматический цикл выполняется
	ELSIF GVL_CELL_CONTROL.xGlobalError THEN
		GVL_HMI.uiPointEditorRejectReason := UINT#7; // Глобальная ошибка
	ELSIF GVL_ROBOT.Status.xBusy OR xPointCheckActive THEN
		GVL_HMI.uiPointEditorRejectReason := UINT#8; // Робот занят
	ELSIF xMotionBusy THEN
		GVL_HMI.uiPointEditorRejectReason := UINT#9; // Motion занят
	ELSIF xDriveError OR GVL_MOTION_MANAGER.stMotionManager.Status.xError THEN
		GVL_HMI.uiPointEditorRejectReason := UINT#10; // Ошибка оси или группы
	ELSIF NOT xPointEditorAllHomed THEN
		GVL_HMI.uiPointEditorRejectReason := UINT#11; // Не выполнен Home
	ELSIF NOT GVL_AXIS_GROUP.AxisGroup.Status.xPositionValid THEN
		GVL_HMI.uiPointEditorRejectReason := UINT#12; // Недостоверные координаты
	ELSIF ((GVL_HMI.uiPointEditorCommand = UINT#2) OR (GVL_HMI.uiPointEditorCommand = UINT#4))
	AND (NOT GVL_POINT_MANAGER.PointManager.Diag.xXLimitValid
		OR NOT GVL_POINT_MANAGER.PointManager.Diag.xYLimitValid
		OR NOT GVL_POINT_MANAGER.PointManager.Diag.xZLimitValid) THEN
		GVL_HMI.uiPointEditorRejectReason := UINT#13; // Software limits недоступны
	END_IF;

	IF (GVL_HMI.uiPointEditorRejectReason = UINT#0) AND (uiPointEditorMagazine <> UINT#0) THEN
		IF (GVL_HMI.uiPointEditorCalibrationMethod <> Persistent_Value.astMagazineCalibration[uiPointEditorMagazine].uiMethod)
		OR ((uiPointEditorReference <> UINT#0) AND (Persistent_Value.astMagazineCalibration[uiPointEditorMagazine].uiMethod <> UINT#3)) THEN
			GVL_HMI.uiPointEditorRejectReason := UINT#25;
		END_IF;
	END_IF;

	IF GVL_HMI.uiPointEditorRejectReason = UINT#0 THEN
		IF GVL_HMI.uiPointEditorCommand = UINT#4 THEN
			InvalidateMagazineCalibration(uiMagazine := uiPointEditorMagazine);
			GVL_HMI.stPointEditorResultPoint := GVL_POINT.Points[ePointEditorName];
			GVL_HMI.uiPointEditorResult := UINT#1;
		ELSIF GVL_HMI.uiPointEditorCommand = UINT#1 THEN
			// CAPTURE возвращает согласованный снимок одного PLC-цикла и не пишет Persistent.
			GVL_HMI.stPointEditorResultPoint.Name := '';
			GVL_HMI.stPointEditorResultPoint.X := GVL_AXIS_GROUP.AxisGroup.Status.ActualX;
			GVL_HMI.stPointEditorResultPoint.Y := GVL_AXIS_GROUP.AxisGroup.Status.ActualY;
			GVL_HMI.stPointEditorResultPoint.Z := GVL_AXIS_GROUP.AxisGroup.Status.ActualZ;
			GVL_HMI.stPointEditorResultPoint.MagazineSafeZ :=
				GVL_HMI.lrPointEditorDraftMagazineSafeZ;
			GVL_HMI.stPointEditorResultPoint.MagazineChangeZ :=
				GVL_HMI.lrPointEditorDraftMagazineChangeZ;
			GVL_HMI.stPointEditorResultPoint.SpeedFactor :=
				GVL_HMI.lrPointEditorDraftSpeedFactor;
			GVL_HMI.stPointEditorResultPoint.xConfigured := FALSE;
			GVL_HMI.uiPointEditorResult := UINT#1;
		ELSIF GVL_HMI.uiPointEditorCommand = UINT#3 THEN
			// CHECK никогда не сохраняет черновик. Сравнение защищает подтверждение
			// на телефоне от изменения точки другим редактором до запуска.
			IF NOT GVL_POINT.Points[ePointEditorName].xConfigured THEN
				GVL_HMI.uiPointEditorRejectReason := UINT#16;
			ELSIF (GVL_POINT.Points[ePointEditorName].X <> GVL_HMI.alrPointEditorDraftXYZ[1])
			OR (GVL_POINT.Points[ePointEditorName].Y <> GVL_HMI.alrPointEditorDraftXYZ[2])
			OR (GVL_POINT.Points[ePointEditorName].Z <> GVL_HMI.alrPointEditorDraftXYZ[3])
			OR (GVL_POINT.Points[ePointEditorName].SpeedFactor <> GVL_HMI.lrPointEditorDraftSpeedFactor)
			OR ((xPointEditorMagazinePoint OR (uiPointEditorGeometryStation <> UINT#0))
				AND ((GVL_POINT.Points[ePointEditorName].MagazineSafeZ <>
					GVL_HMI.lrPointEditorDraftMagazineSafeZ)
				OR (GVL_POINT.Points[ePointEditorName].MagazineChangeZ <>
					GVL_HMI.lrPointEditorDraftMagazineChangeZ))) THEN
				GVL_HMI.uiPointEditorRejectReason := UINT#21;
			ELSE
				xPointCheckRequest := TRUE; // Финальное разрешение после RunMotion/RunCellControl
			END_IF;
		ELSE
			xPointEditorDraftValid :=
				(GVL_HMI.alrPointEditorDraftXYZ[1] >= alrRobotSoftwareMinPosition[1])
				AND (GVL_HMI.alrPointEditorDraftXYZ[1] <= alrRobotSoftwareMaxPosition[1])
				AND (GVL_HMI.alrPointEditorDraftXYZ[2] >= alrRobotSoftwareMinPosition[2])
				AND (GVL_HMI.alrPointEditorDraftXYZ[2] <= alrRobotSoftwareMaxPosition[2])
				AND (GVL_HMI.alrPointEditorDraftXYZ[3] >= alrRobotSoftwareMinPosition[3])
				AND (GVL_HMI.alrPointEditorDraftXYZ[3] <= alrRobotSoftwareMaxPosition[3]);
			IF NOT xPointEditorDraftValid THEN
				GVL_HMI.uiPointEditorRejectReason := UINT#14; // XYZ вне software limits
			ELSIF NOT (((GVL_HMI.lrPointEditorDraftSpeedFactor > 0.1)
				OR ((uiPointEditorGeometryStation <> UINT#0) AND (GVL_HMI.lrPointEditorDraftSpeedFactor >= 0.1)))
			AND (GVL_HMI.lrPointEditorDraftSpeedFactor <= 1.0)) THEN
				GVL_HMI.uiPointEditorRejectReason := UINT#15; // Недопустимая скорость
			ELSIF xPointEditorMagazinePoint
			AND ((GVL_HMI.lrPointEditorDraftMagazineSafeZ < -LREAL#10000.0)
				OR (GVL_HMI.lrPointEditorDraftMagazineSafeZ > LREAL#10000.0)
				OR (GVL_HMI.lrPointEditorDraftMagazineChangeZ < -LREAL#10000.0)
				OR (GVL_HMI.lrPointEditorDraftMagazineChangeZ > LREAL#10000.0)) THEN
				GVL_HMI.uiPointEditorRejectReason := UINT#22; // Смещения магазина вне диапазона
			ELSIF (uiPointEditorGeometryStation <> UINT#0)
			AND NOT ((GVL_HMI.lrPointEditorDraftMagazineSafeZ < LREAL#0.0)
				AND (GVL_HMI.lrPointEditorDraftMagazineSafeZ >= -LREAL#10000.0)
				AND ((GVL_HMI.alrPointEditorDraftXYZ[3] + GVL_HMI.lrPointEditorDraftMagazineSafeZ) >= alrRobotSoftwareMinPosition[3])
				AND ((GVL_HMI.alrPointEditorDraftXYZ[3] + GVL_HMI.lrPointEditorDraftMagazineSafeZ) <= alrRobotSoftwareMaxPosition[3])) THEN
				GVL_HMI.uiPointEditorRejectReason := UINT#22; // SAFE_Z ГК должен поднимать робот в пределах оси
			ELSIF uiPointEditorGeometryStation <> UINT#0 THEN
				// Единственный владелец базы ГК: действующая конфигурация NORMAL/SIMULATION.
				stGeometryConfig.lrX := GVL_HMI.alrPointEditorDraftXYZ[1];
				stGeometryConfig.lrY := GVL_HMI.alrPointEditorDraftXYZ[2];
				stGeometryConfig.lrZ := GVL_HMI.alrPointEditorDraftXYZ[3];
				stGeometryConfig.lrSafeZ := GVL_HMI.lrPointEditorDraftMagazineSafeZ;
				stGeometryConfig.lrChangeZ := stGeometryConfig.lrSafeZ; // Совместимый legacy-канал, отдельного CHANGE нет
				stGeometryConfig.lrSpeedFactor := GVL_HMI.lrPointEditorDraftSpeedFactor;
				stGeometryConfig.xConfigured := TRUE;
				IF GVL_CELL_SETTINGS.eTestEnvironment = E_CELL_TEST_ENVIRONMENT.NORMAL THEN
					Persistent_Value.astConfig[uiPointEditorGeometryStation] := stGeometryConfig;
				ELSE
					Persistent_Value.astSimulationConfig[uiPointEditorGeometryStation] := stGeometryConfig;
				END_IF;
				GVL_GEOMETRY_CONTROL.astActiveConfig[uiPointEditorGeometryStation] := stGeometryConfig;
				GVL_HMI.stPointEditorResultPoint.Name := '';
				GVL_HMI.stPointEditorResultPoint.X := stGeometryConfig.lrX;
				GVL_HMI.stPointEditorResultPoint.Y := stGeometryConfig.lrY;
				GVL_HMI.stPointEditorResultPoint.Z := stGeometryConfig.lrZ;
				GVL_HMI.stPointEditorResultPoint.MagazineSafeZ := stGeometryConfig.lrSafeZ;
				GVL_HMI.stPointEditorResultPoint.MagazineChangeZ := LREAL#0.0;
				GVL_HMI.stPointEditorResultPoint.SpeedFactor := stGeometryConfig.lrSpeedFactor;
				GVL_HMI.stPointEditorResultPoint.xConfigured := TRUE;
				GVL_HMI.uiPointEditorResult := UINT#1;
			ELSIF uiPointEditorReference <> UINT#0 THEN
				stMagazineReferenceDraft.Name := '';
				stMagazineReferenceDraft.X := GVL_HMI.alrPointEditorDraftXYZ[1];
				stMagazineReferenceDraft.Y := GVL_HMI.alrPointEditorDraftXYZ[2];
				stMagazineReferenceDraft.Z := GVL_HMI.alrPointEditorDraftXYZ[3];
				stMagazineReferenceDraft.MagazineSafeZ := 0.0;
				stMagazineReferenceDraft.MagazineChangeZ := 0.0;
				stMagazineReferenceDraft.SpeedFactor := GVL_HMI.lrPointEditorDraftSpeedFactor;
				stMagazineReferenceDraft.xConfigured := TRUE;
				Persistent_Value.astMagazineCalibration[uiPointEditorMagazine].astReference[uiPointEditorReference] := stMagazineReferenceDraft;
				GVL_POINT.Points[ePointEditorName] := stMagazineReferenceDraft;
				GVL_HMI.stPointEditorResultPoint := stMagazineReferenceDraft;
				GVL_HMI.uiPointEditorResult := UINT#1;
			ELSE
				Persistent_Value.astRetainPoints[uiPointStorageIndex].Name := '';
				Persistent_Value.astRetainPoints[uiPointStorageIndex].X :=
					GVL_HMI.alrPointEditorDraftXYZ[1];
				Persistent_Value.astRetainPoints[uiPointStorageIndex].Y :=
					GVL_HMI.alrPointEditorDraftXYZ[2];
				Persistent_Value.astRetainPoints[uiPointStorageIndex].Z :=
					GVL_HMI.alrPointEditorDraftXYZ[3];
				IF xPointEditorMagazinePoint THEN
					Persistent_Value.astRetainPoints[uiPointStorageIndex].MagazineSafeZ :=
						GVL_HMI.lrPointEditorDraftMagazineSafeZ;
					Persistent_Value.astRetainPoints[uiPointStorageIndex].MagazineChangeZ :=
						GVL_HMI.lrPointEditorDraftMagazineChangeZ;
				ELSE
					Persistent_Value.astRetainPoints[uiPointStorageIndex].MagazineSafeZ := LREAL#0.0;
					Persistent_Value.astRetainPoints[uiPointStorageIndex].MagazineChangeZ := LREAL#0.0;
				END_IF;
				Persistent_Value.astRetainPoints[uiPointStorageIndex].SpeedFactor :=
					GVL_HMI.lrPointEditorDraftSpeedFactor;
				Persistent_Value.astRetainPoints[uiPointStorageIndex].xConfigured :=
					NOT xPointEditorMagazinePoint
					OR ((GVL_HMI.lrPointEditorDraftMagazineSafeZ <> LREAL#0.0)
						AND (GVL_HMI.lrPointEditorDraftMagazineChangeZ <> LREAL#0.0));
				GVL_POINT.Points[ePointEditorName] :=
					Persistent_Value.astRetainPoints[uiPointStorageIndex];
				GVL_HMI.stPointEditorResultPoint := GVL_POINT.Points[ePointEditorName];
				GVL_HMI.uiPointEditorResult := UINT#1;
			END_IF;
		END_IF;
	END_IF;

	IF (GVL_HMI.uiPointEditorResult <> UINT#1) AND NOT xPointCheckRequest THEN
		IF GVL_HMI.uiPointEditorCommand = UINT#3 THEN
			uiRobotInterfaceWarningCode := WRN_POINT_CHECK_REJECTED;
		ELSE
			uiRobotInterfaceWarningCode := WRN_POINT_EDIT_REJECTED;
		END_IF;
	END_IF;
	// Ack подтверждает обработку конкретной транзакции даже при отказе.
	IF NOT xPointCheckRequest THEN
		GVL_HMI.udiPointEditorAckSeq := GVL_HMI.udiPointEditorCommandSeq;
	END_IF;
END_IF;

// Плоский OPC UA-интерфейс HMI преобразуется в типизированные запросы FB.
FOR uiMachine := 1 TO 3 DO
	astMachineFaultRequest[uiMachine].xEnabled := GVL_CELL_SETTINGS.xErrorSimulationEnabled;
	astMachineFaultRequest[uiMachine].xReset := GVL_HMI.axMachineSimReset[uiMachine];
	astMachineFaultRequest[uiMachine].xMachineAlarm := GVL_HMI.axMachineSimAlarm[uiMachine];
	astMachineFaultRequest[uiMachine].xDoorFault := GVL_HMI.axMachineSimDoorFault[uiMachine];
	astMachineFaultRequest[uiMachine].xChuckFault := GVL_HMI.axMachineSimChuckFault[uiMachine];
	astMachineFaultRequest[uiMachine].xTimeoutRobotMove := GVL_HMI.axMachineTimeoutRobotMove[uiMachine];
	astMachineFaultRequest[uiMachine].xTimeoutRobotAction := GVL_HMI.axMachineTimeoutRobotAction[uiMachine];
	astMachineFaultRequest[uiMachine].xTimeoutRobotRelease := GVL_HMI.axMachineTimeoutRobotRelease[uiMachine];
	astMachineFaultRequest[uiMachine].xTimeoutDoorOpen := GVL_HMI.axMachineTimeoutDoorOpen[uiMachine];
	astMachineFaultRequest[uiMachine].xTimeoutDoorClose := GVL_HMI.axMachineTimeoutDoorClose[uiMachine];
	astMachineFaultRequest[uiMachine].xTimeoutHatchUnlock := GVL_HMI.axMachineTimeoutHatchUnlock[uiMachine];
	astMachineFaultRequest[uiMachine].xTimeoutChuckOpen := GVL_HMI.axMachineTimeoutChuckOpen[uiMachine];
	astMachineFaultRequest[uiMachine].xTimeoutChuckClose := GVL_HMI.axMachineTimeoutChuckClose[uiMachine];
	astMachineFaultRequest[uiMachine].xTimeoutCycleStart := GVL_HMI.axMachineTimeoutCycleStart[uiMachine];

	astAxisFaultRequest[uiMachine].xEnabled := GVL_CELL_SETTINGS.xErrorSimulationEnabled;
	astAxisFaultRequest[uiMachine].xJogConflict := GVL_HMI.axSimAxisJogConflict[uiMachine];
END_FOR;

stAxisGroupFaultRequest.xEnabled := GVL_CELL_SETTINGS.xErrorSimulationEnabled;
stAxisGroupFaultRequest.xExecute := GVL_HMI.xSimAxisGroupError;

stRobotFaultRequest.xEnabled := GVL_CELL_SETTINGS.xErrorSimulationEnabled;
stRobotFaultRequest.xWrongAction := GVL_HMI.xSimRobotWrongAction;
stRobotFaultRequest.stGripper.xEnabled := GVL_CELL_SETTINGS.xErrorSimulationEnabled;
stRobotFaultRequest.stGripper.xGripper1Fault := GVL_HMI.xSimGripper1Fault;
stRobotFaultRequest.stGripper.xGripper2Fault := GVL_HMI.xSimGripper2Fault;
stRobotFaultRequest.stGripper.xRotationFault := GVL_HMI.xSimGripperRotationFault;
stRobotFaultRequest.stGripper.xGlobalFault := GVL_HMI.xSimGripperGlobalFault;

stRobotFaultRequest.stPoint.xEnabled := GVL_CELL_SETTINGS.xErrorSimulationEnabled;
stRobotFaultRequest.stPoint.xXOutOfLimit := GVL_HMI.xSimPointXOutOfLimit;
stRobotFaultRequest.stPoint.xYOutOfLimit := GVL_HMI.xSimPointYOutOfLimit;
stRobotFaultRequest.stPoint.xZOutOfLimit := GVL_HMI.xSimPointZOutOfLimit;
stRobotFaultRequest.stPoint.xInvalidVelocity := GVL_HMI.xSimPointInvalidVelocity;

IF NOT GVL_CELL_SETTINGS.xErrorSimulationEnabled THEN
	adwTestMagazineFaultMask[1] := DWORD#0;
	adwTestMagazineFaultMask[2] := DWORD#0;
END_IF;
astMagazineFaultRequest[1].xEnabled := GVL_CELL_SETTINGS.xErrorSimulationEnabled;
astMagazineFaultRequest[1].xWrongOperation := GVL_HMI.xSimMagazineWrongOperation
	OR ((adwTestMagazineFaultMask[1] AND DWORD#16#0000_0001) <> DWORD#0);
astMagazineFaultRequest[1].xNoBlank := GVL_HMI.xSimMagazineNoBlank
	OR ((adwTestMagazineFaultMask[1] AND DWORD#16#0000_0002) <> DWORD#0);
astMagazineFaultRequest[1].xNoFreeSlot := GVL_HMI.xSimMagazineNoFreeSlot
	OR ((adwTestMagazineFaultMask[1] AND DWORD#16#0000_0004) <> DWORD#0);
astMagazineFaultRequest[1].xInvalidSlot := GVL_HMI.xSimMagazineInvalidSlot
	OR ((adwTestMagazineFaultMask[1] AND DWORD#16#0000_0008) <> DWORD#0);
astMagazineFaultRequest[1].xSlotContent := GVL_HMI.xSimMagazineSlotContent
	OR ((adwTestMagazineFaultMask[1] AND DWORD#16#0000_0010) <> DWORD#0);
astMagazineFaultRequest[1].xGeometry := GVL_HMI.xSimMagazineGeometry
	OR ((adwTestMagazineFaultMask[1] AND DWORD#16#0000_0020) <> DWORD#0);
astMagazineFaultRequest[2].xEnabled := GVL_CELL_SETTINGS.xErrorSimulationEnabled
	AND (adwTestMagazineFaultMask[2] <> DWORD#0);
astMagazineFaultRequest[2].xWrongOperation :=
	(adwTestMagazineFaultMask[2] AND DWORD#16#0000_0001) <> DWORD#0;
astMagazineFaultRequest[2].xNoBlank :=
	(adwTestMagazineFaultMask[2] AND DWORD#16#0000_0002) <> DWORD#0;
astMagazineFaultRequest[2].xNoFreeSlot :=
	(adwTestMagazineFaultMask[2] AND DWORD#16#0000_0004) <> DWORD#0;
astMagazineFaultRequest[2].xInvalidSlot :=
	(adwTestMagazineFaultMask[2] AND DWORD#16#0000_0008) <> DWORD#0;
astMagazineFaultRequest[2].xSlotContent :=
	(adwTestMagazineFaultMask[2] AND DWORD#16#0000_0010) <> DWORD#0;
astMagazineFaultRequest[2].xGeometry :=
	(adwTestMagazineFaultMask[2] AND DWORD#16#0000_0020) <> DWORD#0;

stCellFaultRequest.xEnabled := GVL_CELL_SETTINGS.xErrorSimulationEnabled;
stCellFaultRequest.xBothGrippers := GVL_HMI.xSimCellBothGrippers;

stSafetyFaultRequest.xEnabled := GVL_CELL_SETTINGS.xErrorSimulationEnabled;
FOR uiMachine := UINT#1 TO UINT#4 DO
	stSafetyFaultRequest.axEmergencyStopStation[uiMachine] :=
		GVL_HMI.axSimSafetyEmergencyStopStation[uiMachine];
	stSafetyFaultRequest.axDoorUnlocked[uiMachine] :=
		GVL_HMI.axSimSafetyDoorUnlocked[uiMachine];
END_FOR;
FOR uiMachine := UINT#1 TO UINT#2 DO
	stSafetyFaultRequest.axEmergencyStopCabinet[uiMachine] :=
		GVL_HMI.axSimSafetyEmergencyStopCabinet[uiMachine];
END_FOR;
stSafetyFaultRequest.xEmergencyStopMpg := GVL_HMI.xSimSafetyEmergencyStopMpg;
stSafetyFaultRequest.xPhaseRelayFault := GVL_HMI.xSimSafetyPhaseRelayFault;
stSafetyFaultRequest.xPressureRelayFault := GVL_HMI.xSimSafetyPressureRelayFault;
stSafetyFaultRequest.xSafetyRelayFault := GVL_HMI.xSimSafetyRelayFault;

(* ---- PLC_PRG.ReadIoEmergencyStop.st ---- *)
METHOD PRIVATE ReadIoEmergencyStop

// --- BEGIN IMPLEMENTATION ---

// Отдельный канал: останов не ждёт текущую транзакцию подмены I/O.
xIoEmergencyResetRequested := FALSE;
xIoEmergencyResetRejected := FALSE;
udiIoEmergencyRequestSeq := GVL_HMI.udiIoEmergencyCommandSeq;
IF xIoInitialized AND (udiIoEmergencyRequestSeq <> GVL_HMI.udiIoEmergencyAckSeq) THEN
    IF GVL_HMI.uiIoEmergencyAction = UINT#1 THEN
        xIoManualActive := FALSE;
        GVL_HMI.xIoEmergencyStopActive := TRUE;
        GVL_HMI.uiIoEmergencyResult := UINT#1;
        GVL_HMI.udiIoEmergencyAckSeq := udiIoEmergencyRequestSeq;
    ELSE
        xIoEmergencyResetRequested := TRUE;
    END_IF;
END_IF;
IF GVL_HMI.xIoEmergencyStopActive THEN
    GVL_CELL_CONTROL.xStop := TRUE;
    GVL_CELL_CONTROL.xStart := FALSE;
    GVL_CELL_CONTROL.xEnable := FALSE;
    GVL_CELL_CONTROL.xManual := TRUE;
    GVL_ROBOT.Command.xExecute := FALSE;
    GVL_ROBOT.Command.xStop := TRUE;
    GVL_ROBOT.ModbusCommand.xExecute := FALSE;
    GVL_ROBOT.ModbusCommand.xStop := TRUE;
    GVL_HMI.xRobotManualExecute := FALSE;
    GVL_HMI.stRobotCommand.xExecute := FALSE;
    xPointCheckStopRequest := xPointCheckActive;
    FOR uiIoIndex := UINT#1 TO UINT#3 DO
        GVL_HMI.astAxisHmiCommand[uiIoIndex].xJogPositive := FALSE;
        GVL_HMI.astAxisHmiCommand[uiIoIndex].xJogNegative := FALSE;
        GVL_HMI.astAxisHmiCommand[uiIoIndex].xHome := FALSE;
        GVL_HMI.astAxisHmiCommand[uiIoIndex].xMoveAbsolute := FALSE;
        GVL_HMI.astAxisHmiCommand[uiIoIndex].xMoveRelative := FALSE;
        GVL_HMI.axMachineManualHatchOpen[uiIoIndex] := FALSE;
        GVL_HMI.axMachineManualHatchClose[uiIoIndex] := FALSE;
        GVL_HMI.axMachineManualHatchUnlock[uiIoIndex] := FALSE;
        GVL_HMI.axMachineManualHatchLock[uiIoIndex] := FALSE;
        GVL_HMI.axMachineManualChuckOpen[uiIoIndex] := FALSE;
        GVL_HMI.axMachineManualChuckClose[uiIoIndex] := FALSE;
    END_FOR;
END_IF;
